// TwinCAT 3 PLC project Untitled1
// ProgramVersion: 3.1.4024.0
// libraries:
//   CmpBitmapPool, * (System)
//   Tc2_ControllerToolbox, * (Beckhoff Automation GmbH)
//   Tc2_MC2, * (Beckhoff Automation GmbH)
//   Tc2_Standard, * (Beckhoff Automation GmbH)
//   Tc2_System, * (Beckhoff Automation GmbH)
//   Tc2_Utilities, * (Beckhoff Automation GmbH)
//   Tc3_Module, * (Beckhoff Automation GmbH)
//   VisuSymbols,3.5.10.0,System
// project tree:
//   DUTs/Cartesian Space/ ST_CartesianAdditionalParametes.TcDUT, ST_CartesianForces.TcDUT, ST_CartesianPose.TcDUT, ST_CartesianState.TcDUT, ST_CartesianTarget.TcDUT, ST_CartesianVelocity.TcDUT
//   DUTs/ En_TargetMode.TcDUT, E_CalibrationState.TcDUT, E_ControllerType.TcDUT, E_GameID.TcDUT, E_Language.TcDUT, E_MainState.TcDUT, E_RehabMode.TcDUT, ST_HomingResult.TcDUT, ST_TherapyConfig.TcDUT
//   DUTs/Joint Space/ ST_JointPose.TcDUT, ST_JointState.TcDUT, ST_JointTarget.TcDUT, ST_JointTorque.TcDUT, ST_JointVelocity.TcDUT
//   / GlobalTextList.TcGTLO, PlcTask.TcTTO, Visualization Manager.TcVMO (not stored)
//   GVLs/ GVL_ConstantCoefficent.TcGVL, GVL_AbsoluteEncoders.TcGVL, GVL_Axes.TcGVL, GVL_Current.TcGVL, GVL_EndeffectorPosition.TcGVL, GVL_ForceTorqueSensor.TcGVL, GVL_GamePong.TcGVL, GVL_HMI.TcGVL, GVL_HomingResult.TcGVL, GVL_MessageStaus.TcGVL, GVL_MicroSwitch.TcGVL, GVL_RobotData.TcGVL, GVL_StatusAxes.TcGVL, GVL_TargetPoints.TcGVL, GVL_Torque.TcGVL
//   POUs/Crazy Car/ FB_CrazyCarGame.TcPOU, ST_CrazyCarToUnity.TcDUT, ST_UnityToCrazyCar.TcDUT
//   POUs/ FB_AdmittanceController.TcPOU, FB_DoHoming.TcPOU, FB_DriveInterface.TcPOU, FB_DynamicsCompensator.TcPOU, FB_ForceController.TcPOU, FB_ForceTorqueSensor.TcPOU, FB_ImpedanceController.TcPOU, FB_LanguageManager.TcPOU, FB_LaunchGame.TcPOU, FB_RobotIsActive.TcPOU, FB_StartGame.TcPOU, FB_SwitchOpMode.TcPOU, FB_TherapyManager.TcPOU, FB_ThreeAxisSafety.TcPOU, FB_RobotKinematics.TcPOU, HardwareWallCheck.TcPOU, MAIN.TcPOU, FB_JointStateReader.TcPOU, FB_VirtuallWall.TcPOU, StopAllMotion.TcPOU
//   POUs/Firrfly Game/ FB_FireflyGame.TcPOU, ST_FireflyFromUnity.TcDUT, ST_FireflyToUnity.TcDUT
//   POUs/HMI_FunBlock/ FB_HMI_Monitoring.TcPOU, FB_HMI_TherapyConfiguration.TcPOU, FB_UserSecuring.TcPOU, MicroswitchCheck.TcPOU
//   POUs/PeelerGame/ ST_PeelerFromUnity.TcDUT, FB_PeelingGame.TcPOU, ST_PeelerToUnity.TcDUT
//   POUs/Sorter Game/ FB_SorterGame.TcPOU, ST_SorterToUnity.TcDUT, ST_UnityToSorter.TcDUT
//   VISUs/ ImagePool.TcIPO (not stored), Screen2.TcVIS, Visualization.TcVIS
// real-time tasks:
//   TASK PlcTask: cycle T#10ms, priority 20, ADS port 350
//   TASK VISU_TASK1: cycle T#200000us, priority 1, ADS port 352
// motion (NC):
//   TASK NC-Task 1 SAF: cycle T#1ms, priority 4, ADS port 501
//   TASK NC-Task 1 SVB: cycle T#1ms, priority 6, ADS port 511
//   AXIS Motor-A (id 1)
//     Velo: Maximum=80
//     OtherSettings: AllowMotionCmdToSlave=true
//     encoder EncType=19
//       EncPara: MaxCount=#xffffffff
//         TimeComp: TimeCompMode=1
//     drive DrvType=16
//       DrvPara: MaxCount=#xffffffff, DriveControlDWord=#x00020000
//         Analog: TorqueSetpointScale=10, ScaleFactorActTorque=0.1
//         TimeComp: TaskDelayCycles=1
//     controller CtrType=1
//       CtrPara: PriorControlFactor=1
//         PosDiffControl: Enable=false
//         Observer: BandWidth=20
//   AXIS Motor-B (id 3)
//     Velo: Maximum=80
//     OtherSettings: AllowMotionCmdToSlave=true
//     encoder EncType=19
//       EncPara: MaxCount=#xffffffff
//         TimeComp: TimeCompMode=1
//     drive DrvType=16
//       DrvPara: MaxCount=#xffffffff, DriveControlDWord=#x00020000
//         Analog: TorqueSetpointScale=10, ScaleFactorActTorque=0.1
//         TimeComp: TaskDelayCycles=1
//     controller CtrType=1
//       CtrPara: PriorControlFactor=1
//         PosDiffControl: Enable=false, Range=20
//         Observer: BandWidth=20
//   AXIS Motor-C (id 2)
//     Velo: Maximum=80
//     OtherSettings: AllowMotionCmdToSlave=true
//     encoder EncType=19
//       EncPara: MaxCount=#xffffffff
//         TimeComp: TimeCompMode=1
//     drive DrvType=16
//       DrvPara: MaxCount=#xffffffff, DriveControlDWord=#x00020000
//         Analog: TorqueSetpointScale=10, ScaleFactorActTorque=0.1
//         TimeComp: TaskDelayCycles=1
//     controller CtrType=1
//       CtrPara: PriorControlFactor=1
//         PosDiffControl: Enable=false
//         Observer: BandWidth=20
// I/O:
//   DEVICE Device 3 (EtherCAT), AmsNetId 10.4.37.185.4.1
//     Motor-A [EPOS4 Module 50/8 EtherCAT]
//       modules: Module 1 (CSP Mode)
//     Motor-B [EPOS4 Module 50/8 EtherCAT]
//       modules: Module 1 (CSP Mode)
//     Motor-C [EPOS4 Module 50/8 EtherCAT]
//       modules: Module 1 (CSP Mode)
//     Box 7 (RFT_EC02) [RFT_EC02]
// variable links:
//   NC-Task 1 SAF/Axes/Motor-A <-> Device 3 (EtherCAT)/Motor-A
//     Drive/Inputs/In/nDataIn3[0] <-> Module 1 (CSP Mode)/CSP Inputs/Torque actual value
//     Drive/Inputs/In/nDcOutputTime <-> InfoData/DcOutputShift
//     Drive/Inputs/In/nState1 <-> Module 1 (CSP Mode)/CSP Inputs/Statusword
//     Drive/Inputs/In/nState2 <-> Module 1 (CSP Mode)/CSP Inputs/Statusword @bit 8
//     Drive/Inputs/In/nState4 @bit 1 <-> WcState/InputToggle
//     Drive/Inputs/In/nState4 <-> WcState/WcState
//     Drive/Inputs/In/nState5 <-> Module 1 (CSP Mode)/CSP Inputs/Mode of operation display
//     Drive/Outputs/Out/nCtrl1 <-> Module 1 (CSP Mode)/CSP Outputs/Controlword
//     Drive/Outputs/Out/nCtrl2 <-> Module 1 (CSP Mode)/CSP Outputs/Controlword @bit 8
//     Drive/Outputs/Out/nCtrl5 <-> Module 1 (CSP Mode)/CSP Outputs/Mode of operation
//     Drive/Outputs/Out/nDataOut1 <-> Module 1 (CSP Mode)/CSP Outputs/Target position
//     Drive/Outputs/Out/nDataOut2 <-> Module 1 (CSP Mode)/CSP Outputs/Target velocity
//     Drive/Outputs/Out/nDataOut3[0] <-> Module 1 (CSP Mode)/CSP Outputs/Torque offset
//     Drive/Outputs/Out/nDataOut4[0] <-> Module 1 (CSP Mode)/CSP Outputs/Target torque
//     Enc/Inputs/In/nDataIn1 <-> Module 1 (CSP Mode)/CSP Inputs/Position actual value
//     Enc/Inputs/In/nDataIn7 <-> Module 1 (CSP Mode)/CSP Inputs/Velocity actual value
//     Enc/Inputs/In/nDcInputTime <-> InfoData/DcInputShift
//     Enc/Inputs/In/nState4 @bit 1 <-> WcState/InputToggle
//     Enc/Inputs/In/nState4 <-> WcState/WcState
//   NC-Task 1 SAF/Axes/Motor-B <-> Device 3 (EtherCAT)/Motor-B
//     Drive/Inputs/In/nDataIn3[0] <-> Module 1 (CSP Mode)/CSP Inputs/Torque actual value
//     Drive/Inputs/In/nDcOutputTime <-> InfoData/DcOutputShift
//     Drive/Inputs/In/nState1 <-> Module 1 (CSP Mode)/CSP Inputs/Statusword
//     Drive/Inputs/In/nState2 <-> Module 1 (CSP Mode)/CSP Inputs/Statusword @bit 8
//     Drive/Inputs/In/nState4 @bit 1 <-> WcState/InputToggle
//     Drive/Inputs/In/nState4 <-> WcState/WcState
//     Drive/Inputs/In/nState5 <-> Module 1 (CSP Mode)/CSP Inputs/Mode of operation display
//     Drive/Outputs/Out/nCtrl1 <-> Module 1 (CSP Mode)/CSP Outputs/Controlword
//     Drive/Outputs/Out/nCtrl2 <-> Module 1 (CSP Mode)/CSP Outputs/Controlword @bit 8
//     Drive/Outputs/Out/nCtrl5 <-> Module 1 (CSP Mode)/CSP Outputs/Mode of operation
//     Drive/Outputs/Out/nDataOut1 <-> Module 1 (CSP Mode)/CSP Outputs/Target position
//     Drive/Outputs/Out/nDataOut2 <-> Module 1 (CSP Mode)/CSP Outputs/Target velocity
//     Drive/Outputs/Out/nDataOut3[0] <-> Module 1 (CSP Mode)/CSP Outputs/Torque offset
//     Drive/Outputs/Out/nDataOut4[0] <-> Module 1 (CSP Mode)/CSP Outputs/Target torque
//     Enc/Inputs/In/nDataIn1 <-> Module 1 (CSP Mode)/CSP Inputs/Position actual value
//     Enc/Inputs/In/nDataIn7 <-> Module 1 (CSP Mode)/CSP Inputs/Velocity actual value
//     Enc/Inputs/In/nDcInputTime <-> InfoData/DcInputShift
//     Enc/Inputs/In/nState4 @bit 1 <-> WcState/InputToggle
//     Enc/Inputs/In/nState4 <-> WcState/WcState
//   NC-Task 1 SAF/Axes/Motor-C <-> Device 3 (EtherCAT)/Motor-C
//     Drive/Inputs/In/nDataIn3[0] <-> Module 1 (CSP Mode)/CSP Inputs/Torque actual value
//     Drive/Inputs/In/nDcOutputTime <-> InfoData/DcOutputShift
//     Drive/Inputs/In/nState1 <-> Module 1 (CSP Mode)/CSP Inputs/Statusword
//     Drive/Inputs/In/nState2 <-> Module 1 (CSP Mode)/CSP Inputs/Statusword @bit 8
//     Drive/Inputs/In/nState4 @bit 1 <-> WcState/InputToggle
//     Drive/Inputs/In/nState4 <-> WcState/WcState
//     Drive/Inputs/In/nState5 <-> Module 1 (CSP Mode)/CSP Inputs/Mode of operation display
//     Drive/Outputs/Out/nCtrl1 <-> Module 1 (CSP Mode)/CSP Outputs/Controlword
//     Drive/Outputs/Out/nCtrl2 <-> Module 1 (CSP Mode)/CSP Outputs/Controlword @bit 8
//     Drive/Outputs/Out/nCtrl5 <-> Module 1 (CSP Mode)/CSP Outputs/Mode of operation
//     Drive/Outputs/Out/nDataOut1 <-> Module 1 (CSP Mode)/CSP Outputs/Target position
//     Drive/Outputs/Out/nDataOut2 <-> Module 1 (CSP Mode)/CSP Outputs/Target velocity
//     Drive/Outputs/Out/nDataOut3[0] <-> Module 1 (CSP Mode)/CSP Outputs/Torque offset
//     Drive/Outputs/Out/nDataOut4[0] <-> Module 1 (CSP Mode)/CSP Outputs/Target torque
//     Enc/Inputs/In/nDataIn1 <-> Module 1 (CSP Mode)/CSP Inputs/Position actual value
//     Enc/Inputs/In/nDataIn7 <-> Module 1 (CSP Mode)/CSP Inputs/Velocity actual value
//     Enc/Inputs/In/nDcInputTime <-> InfoData/DcInputShift
//     Enc/Inputs/In/nState4 @bit 1 <-> WcState/InputToggle
//     Enc/Inputs/In/nState4 <-> WcState/WcState
//   Untitled1/Untitled1 Instance <-> Device 3 (EtherCAT)/Box 7 (RFT_EC02)
//     PlcTask Inputs/GVL_ForceTorqueSensor.RawFx <-> IN_GENERIC process data mapping/Raw_Fx
//     PlcTask Inputs/GVL_ForceTorqueSensor.RawFy <-> IN_GENERIC process data mapping/Raw_Fy
//     PlcTask Inputs/GVL_ForceTorqueSensor.RawFz <-> IN_GENERIC process data mapping/Raw_Fz
//     PlcTask Inputs/GVL_ForceTorqueSensor.RawMx <-> IN_GENERIC process data mapping/Raw_Tx
//     PlcTask Inputs/GVL_ForceTorqueSensor.RawMy <-> IN_GENERIC process data mapping/Raw_Ty
//     PlcTask Inputs/GVL_ForceTorqueSensor.RawMz <-> IN_GENERIC process data mapping/Raw_Tz
//     PlcTask Outputs/GVL_ForceTorqueSensor.ConfigParameter <-> OUT_GENERIC process data mapping/ConfigParam_1
//   Untitled1/Untitled1 Instance <-> Device 3 (EtherCAT)/Motor-A
//     PlcTask Inputs/GVL_AbsoluteEncoders.AbsoluteBetaPosition <-> Module 1 (CSP Mode)/CSP Inputs/Position actual value sensor 2
//     PlcTask Inputs/GVL_Current.MotorCurrentM1_mA <-> Module 1 (CSP Mode)/CSP Inputs/Current actual value averaged
//     PlcTask Inputs/GVL_MicroSwitch.dwMicroSwitchDriverA <-> Module 1 (CSP Mode)/CSP Inputs/Digital inputs
//   Untitled1/Untitled1 Instance <-> Device 3 (EtherCAT)/Motor-B
//     PlcTask Inputs/GVL_AbsoluteEncoders.AbsoluteLinearPosition <-> Module 1 (CSP Mode)/CSP Inputs/Position actual value sensor 2
//     PlcTask Inputs/GVL_Current.MotorCurrentM2_mA <-> Module 1 (CSP Mode)/CSP Inputs/Current actual value averaged
//     PlcTask Inputs/GVL_MicroSwitch.dwMicroSwitchDriverB <-> Module 1 (CSP Mode)/CSP Inputs/Digital inputs
//   Untitled1/Untitled1 Instance <-> Device 3 (EtherCAT)/Motor-C
//     PlcTask Inputs/GVL_AbsoluteEncoders.AbsoluteTetaPosition <-> Module 1 (CSP Mode)/CSP Inputs/Position actual value sensor 2
//     PlcTask Inputs/GVL_Current.MotorCurrentM3_mA <-> Module 1 (CSP Mode)/CSP Inputs/Current actual value averaged
//   Untitled1/Untitled1 Instance <-> NC-Task 1 SAF/Axes/Motor-A
//     PlcTask Inputs/GVL_Axes.Axis1.NcToPlc <-> Outputs/ToPlc
//     PlcTask Inputs/GVL_Torque.TorqueM1_Act <-> Outputs/ToPlc/ActTorque
//     PlcTask Outputs/GVL_Axes.Axis1.PlcToNc <-> Inputs/FromPlc
//   Untitled1/Untitled1 Instance <-> NC-Task 1 SAF/Axes/Motor-B
//     PlcTask Inputs/GVL_Axes.Axis2.NcToPlc <-> Outputs/ToPlc
//     PlcTask Inputs/GVL_Torque.TorqueM2_Act <-> Outputs/ToPlc/ActTorque
//     PlcTask Outputs/GVL_Axes.Axis2.PlcToNc <-> Inputs/FromPlc
//   Untitled1/Untitled1 Instance <-> NC-Task 1 SAF/Axes/Motor-C
//     PlcTask Inputs/GVL_Axes.Axis3.NcToPlc <-> Outputs/ToPlc
//     PlcTask Inputs/GVL_Torque.TorqueM3_Act <-> Outputs/ToPlc/ActTorque
//     PlcTask Outputs/GVL_Axes.Axis3.PlcToNc <-> Inputs/FromPlc

CONFIGURATION Untitled1
    RESOURCE PLC ON TwinCAT3
        TASK PlcTask(INTERVAL := T#10ms, PRIORITY := 20);
        PROGRAM MAIN WITH PlcTask : MAIN;
    END_RESOURCE
END_CONFIGURATION

// ---- DUTs/Cartesian Space/ST_CartesianAdditionalParametes.TcDUT
TYPE ST_CartesianAdditionalParametes :
STRUCT
	BetaIncremental : LREAL;
	RIncremental : LREAL;
	X_Dir_Abs :LREAL;
	Y_Dir_Abs :LREAL;
	WristAngle_Abs : LREAL;

END_STRUCT
END_TYPE

// ---- DUTs/Cartesian Space/ST_CartesianForces.TcDUT
TYPE ST_CartesianForces :
STRUCT
	Fx     : LREAL; // Linear force along X (N)
    Fy     : LREAL; // Linear force along Y (N)
    Mtheta : LREAL; // Moment/Torque around Theta wrist axis (Nm)
END_STRUCT
END_TYPE

// ---- DUTs/Cartesian Space/ST_CartesianPose.TcDUT
TYPE ST_CartesianPose :
STRUCT
	X     : LREAL; // X position (mm)
    Y     : LREAL; // Y position (mm)
    Theta : LREAL; // Wrist angle (deg / rad)
END_STRUCT
END_TYPE

// ---- DUTs/Cartesian Space/ST_CartesianState.TcDUT
TYPE ST_CartesianState :
STRUCT
	Position : ST_CartesianPose;     // Contains X, Y, Theta
    Velocity : ST_CartesianVelocity; // Contains Vx, Vy, Vtheta
	Force    : ST_CartesianForces;    // Contains Fx, Fy, Mtheta
END_STRUCT
END_TYPE

// ---- DUTs/Cartesian Space/ST_CartesianTarget.TcDUT
TYPE ST_CartesianTarget :
STRUCT
	Position : ST_CartesianPose;     // Game target position
    Velocity : ST_CartesianVelocity; // Feedforward target velocity
    Force    : ST_CartesianForces;    // Force setpoint (e.g. 0 N for admittance)
END_STRUCT
END_TYPE

// ---- DUTs/Cartesian Space/ST_CartesianVelocity.TcDUT
TYPE ST_CartesianVelocity :
STRUCT
	Vx     : LREAL; // Linear velocity along X (mm/s or m/s)
    Vy     : LREAL; // Linear velocity along Y (mm/s or m/s)
    Vtheta : LREAL; // Angular velocity around Theta (deg/s or rad/s)
END_STRUCT
END_TYPE

// ---- DUTs/En_TargetMode.TcDUT
{attribute 'qualified_only'}
{attribute 'strict'}
TYPE En_TargetMode :
(
	eCSP := 4,   // Cyclic Synchronous Position
    eCSV := 2,   // Cyclic Synchronous Velocity
    eCST := 1   // Cyclic Synchronous Torque
);
END_TYPE

// ---- DUTs/E_CalibrationState.TcDUT
{attribute 'qualified_only'}
{attribute 'strict'}
TYPE E_CalibrationState :
(
	INIT,
    SET_FILTER,
    START,
    WaitingforCalibrationButton,
    ZEROING,
    RUNNING
);
END_TYPE

// ---- DUTs/E_ControllerType.TcDUT
{attribute 'qualified_only'}
{attribute 'strict'}
TYPE E_ControllerType :
(
    ControlNone         := 0,

    ControlPosition     := 1,

    ControlVelocity     := 2,

    ControlTorque       := 3,

    ControlForce        := 4,

    ControlImpedance    := 5,

    ControlAdmittance   := 6,

    ControlHybrid       := 7,

    ControlCustom       := 8
);
END_TYPE

// ---- DUTs/E_GameID.TcDUT
{attribute 'qualified_only'}
{attribute 'strict'}
TYPE E_GameID :
(
    NONE        := 0,
    PONG        := 1,
    PEELING     := 2,
    GOLD_MINER  := 3,
    BALLOON     := 4,
    SNOW_WIPER  := 5,
    SORTER      := 6,
    FLOWER      := 7,
    CRAZY_CAR   := 8
);
END_TYPE

// ---- DUTs/E_Language.TcDUT
{attribute 'qualified_only'}
{attribute 'strict'}
TYPE E_Language :
(
	EN,
    FR
);
END_TYPE

// ---- DUTs/E_MainState.TcDUT
{attribute 'qualified_only'}
{attribute 'strict'}
TYPE E_MainState :
(
	Init                := 0,
    Homing              := 10,
    ClearNCErrors       := 20,
    ChangingDriverMode        := 30,
    Standby             := 40,  // NEW: Motors are ON, holding position, waiting for HMI start
    RunningTherapy      := 50,  // NEW: The robot is actively doing rehab
    Fault               := 99
);
END_TYPE

// ---- DUTs/E_RehabMode.TcDUT
{attribute 'qualified_only'}
{attribute 'strict'}
TYPE E_RehabMode :
(
	ModeIdle              := 0, // Safety default: system is ready but therapy is not active
    ModePassive           := 1, // Robot moves a completely relaxed patient rigidly along a path
    ModeActiveFree        := 2, // Robot is totally transparent; patient moves freely without resistance
    ModeActiveAssistive   := 3, // Robot provides assistive forces to help the patient reach the target
    ModeActiveResistive   := 4, // Robot pushes against the patient to build muscle strength
    ModePerturbation      := 5, // Robot applies sudden, unexpected forces to train patient reflexes
    ModeAssessment        := 6  // Robot measures patient capability passively without providing assistance
);
END_TYPE

// ---- DUTs/Joint Space/ST_JointPose.TcDUT
TYPE ST_JointPose :
STRUCT
	q1 : LREAL;
    q2 : LREAL;
    q3 : LREAL;
END_STRUCT
END_TYPE

// ---- DUTs/Joint Space/ST_JointState.TcDUT
TYPE ST_JointState :
STRUCT
	Position : ST_JointPose; // Current joint angles (J1, J2, J3)
    Velocity : ST_JointVelocity; // Current joint speeds (J1, J2, J3)
    Torque   : ST_JointTorque; // Measured motor torques (J1, J2, J3)
END_STRUCT
END_TYPE

// ---- DUTs/Joint Space/ST_JointTarget.TcDUT
TYPE ST_JointTarget :
STRUCT
	Position : ST_JointPose; // Commanded joint angles
    Velocity : ST_JointVelocity; // Commanded joint speeds
    Torque   : ST_JointTorque; // Calculated motor torques (T1, T2, T3)
END_STRUCT
END_TYPE

// ---- DUTs/Joint Space/ST_JointTorque.TcDUT
TYPE ST_JointTorque :
STRUCT
	M1 : LREAL;
    M2 : LREAL;
    M3 : LREAL;
END_STRUCT
END_TYPE

// ---- DUTs/Joint Space/ST_JointVelocity.TcDUT
TYPE ST_JointVelocity :
STRUCT
	q1_dot : LREAL; // dq1 / dt
    q2_dot : LREAL; // dq2 / dt
    q3_dot : LREAL; // dq3 / dt
END_STRUCT
END_TYPE

// ---- DUTs/ST_HomingResult.TcDUT
TYPE ST_HomingResult :
STRUCT
	HomePos_Beta  : LREAL;   (* joint angle/position after homing *)
    HomePos_Theta  : LREAL;
    HomePos_R  : LREAL;
END_STRUCT
END_TYPE

// ---- DUTs/ST_TherapyConfig.TcDUT
TYPE ST_TherapyConfig :
STRUCT
	// 1. Core Selections
    TherapyMode          : E_RehabMode;
    ControllerType       : E_ControllerType;
    
    // 2. Feature Flags
    FeatureInertiaComp   : BOOL;  
    FeatureFrictionComp  : BOOL; 
    FeatureVirtualWall   : BOOL; 
	
//    FeatureDataLogger    : BOOL; 
    
    // 3. Global Safety Limits (Apply to ALL controllers)
    GlobalForceLimit     : LREAL := 50 ; // Maximum safe force allowed
    GlobalVelocityLimit  : LREAL; // Maximum safe speed allowed (please clarify : is it in Jointspace or Cartesian space)
	
	Stiffness_K         : LREAL; // Virtual spring stiffness for Impedance
    Damping_D           : LREAL; // Virtual friction/viscosity for Impedance
    Mass_M              : LREAL; // Virtual mass for Admittance
END_STRUCT
END_TYPE

// ---- POUs/Crazy Car/ST_CrazyCarToUnity.TcDUT
TYPE ST_CrazyCarToUnity :
STRUCT
	fY           : REAL;   // gas, Y position 0..100 %
    fWristAngle  : REAL;   // wrist angle, degrees, 0 = home
    GameIsActive : BOOL;
END_STRUCT
END_TYPE

// ---- POUs/Crazy Car/ST_UnityToCrazyCar.TcDUT
TYPE ST_UnityToCrazyCar  :
STRUCT
	bGameClosed : BOOL;   // TRUE = Unity game closed
    nGameStatus : INT;    // 0 = menu/popup, 1 = Taxi, 2 = Van, 3 = Truck
END_STRUCT
END_TYPE

// ---- POUs/Firrfly Game/ST_FireflyFromUnity.TcDUT
{attribute 'pack_mode' := '1'}
TYPE ST_FireflyFromUnity :
STRUCT
    nGameStatus  : INT;    // 0 = menu/results, 1/2/3 = playing Level 1/2/3, 4 = paused
    bExitPressed : BOOL;   // TRUE for ~0.2 s when an Exit button is pressed, then FALSE
    bWrongFlower : BOOL;   // TRUE for ~0.2 s each time a wrong flower is selected, then FALSE
END_STRUCT
END_TYPE

// ---- POUs/Firrfly Game/ST_FireflyToUnity.TcDUT
TYPE ST_FireflyToUnity :
STRUCT
    fX : REAL;   // -100..+100 %, 0 = home (middle of the scene), +100 = right edge of the garden
    fY : REAL;   // -100..+100 %, 0 = home (middle of the scene), +100 = top edge (robot forward)
END_STRUCT
END_TYPE

// ---- POUs/PeelerGame/ST_PeelerFromUnity.TcDUT
{attribute 'pack_mode' := '1'}
TYPE ST_PeelerFromUnity :
STRUCT
	bInContact    : BOOL;    // Fruit collision state
    nObjectType   : INT;     // 1 = Kiwi, 2 = Orange, 3 = Pineapple
    bGameFinished : BOOL;    // TRUE when the user clicks the Close button in Unity
END_STRUCT
END_TYPE

// ---- POUs/PeelerGame/ST_PeelerToUnity.TcDUT
TYPE ST_PeelerToUnity :
STRUCT
	fY          : REAL;    // Y position (0 - 100%)
	GameIsActive : BOOL;
   

END_STRUCT
END_TYPE

// ---- POUs/Sorter Game/ST_SorterToUnity.TcDUT
TYPE ST_SorterToUnity :
STRUCT
    fX           : REAL;    // X position 0–100%
    GameIsActive : BOOL;
END_STRUCT
END_TYPE

// ---- POUs/Sorter Game/ST_UnityToSorter.TcDUT
TYPE ST_UnityToSorter :
STRUCT
	bGameClosed : BOOL;   // TRUE = Unity game closed
    nGameStatus : INT;    // 0 = not playing, 1 = light, 2 = medium, 3 = heavy
END_STRUCT
END_TYPE

// ---- GVLs/GVL_ConstantCoefficent.TcGVL
{attribute 'qualified_only'}
// These number is checked two times, the error between Absolute and Incremental Encoder is under 1% that is acceptable
// Root of error is related to timing belt 


VAR_GLOBAL
	K2: LREAL :=24.40;  // calculate with result of absolute encoder
	
	K3: LREAL :=219.726; // calculate with result of absolute encoder
	K1: LREAL := 9.97; // calculate with result of absolute encoder
	
END_VAR

// ---- GVLs/GVL_AbsoluteEncoders.TcGVL
{attribute 'qualified_only'}
VAR_GLOBAL
	AbsoluteBetaPosition AT %I* : DINT;
	AbsoluteLinearPosition AT %I* : DINT;
	AbsoluteTetaPosition AT %I* : DINT;
END_VAR

// ---- GVLs/GVL_Axes.TcGVL
{attribute 'qualified_only'}
VAR_GLOBAL
	Axis1 : AXIS_REF;
	Axis2 : AXIS_REF;
	Axis3 : AXIS_REF;
END_VAR

// ---- GVLs/GVL_Current.TcGVL
{attribute 'qualified_only'}
VAR_GLOBAL
	MotorCurrentM1_mA AT %I* : DINT; // PDO value from EPOS4 [mA]
	MotorCurrentM2_mA AT %I* : DINT;
	MotorCurrentM3_mA AT %I* : DINT;
	MotorCurrentM1_A : LREAL;  // // Converted current [A]
	MotorCurrentM2_A : LREAL;
	MotorCurrentM3_A : LREAL;
	
END_VAR

// ---- GVLs/GVL_EndeffectorPosition.TcGVL
{attribute 'qualified_only'}
VAR_GLOBAL
	WristAngle : LREAL;
	X_Dir : LREAL;
	Y_Dir : LREAL;
	R_Dir : LREAL;
	Beta : LREAL;
	
	X_Dir_Abs: LREAL;
	Y_Dir_Abs: LREAL;
	R_Dir_Abs: LREAL;
	BetaFromAbsolute : LREAL;
	WristAngle_Abs: LREAL;
	
END_VAR

// ---- GVLs/GVL_ForceTorqueSensor.TcGVL
{attribute 'qualified_only'}
VAR_GLOBAL
	ConfigParameter AT %Q* : DWORD;
	RawFx AT %I* : INT;
	RawFy AT %I* : INT;
	RawFz AT %I* : INT;
	RawMx AT %I* : INT;
	RawMy AT %I* : INT;
	RawMz AT %I* : INT;
	
	//
	Fx_ActFTS : LREAL;    // N
	Fy_ActFTS : LREAL;
	Mz_ActFTS : LREAL;    //N.M
	
END_VAR

// ---- GVLs/GVL_GamePong.TcGVL
{attribute 'qualified_only'}
VAR_GLOBAL
	// Robot Position for Unity (0-100)
    MyRobotY : REAL ;
END_VAR

// ---- GVLs/GVL_HMI.TcGVL
{attribute 'qualified_only'}
VAR_GLOBAL
	


	
	bLaunchGameSpongCmd : BOOL := FALSE;
	bLaunchGamePeelerCmd : BOOL := FALSE;
	bLaunchGameGoldMiner : BOOL := FALSE;
	bLaunchGameBalloonAssesment : BOOL := FALSE;
	bLaunchGameSnowWiper : BOOL := FALSE;
	bLaunchGameSorter : BOOL := FALSE;
	bLaunchGameFlower : BOOL := FALSE;
	bLaunchGameCrazyCar : BOOL := FALSE;
	
	
	
	
	
	// MicroSwitch Check
	CheckMicroswitchLinearMin : BOOL := FALSE;
	CheckMicroswitchLinearMax : BOOL := FALSE;
	CheckMicroswitchRotationLeft : BOOL := FALSE;
	CheckMicroswitchRotationRight : BOOL := FALSE;
	CheckMicroswitchWristLeft : BOOL := FALSE;
	CheckMicroswitchWristRight : BOOL := FALSE;
	
	HardwareLimitisActived : BOOL := FALSE;
	
	
			// HMIHardwareMicroSwitch Check for activation
	
	HwCheckMicroswitchLinearMin : BOOL := FALSE;
	HwCheckMicroswitchLinearMax : BOOL := FALSE;
	HwCheckMicroswitchRotationLeft : BOOL := FALSE;
	HwCheckMicroswitchRotationRight : BOOL := FALSE;
	HwCheckMicroswitchWristLeft : BOOL := FALSE;
	HwCheckMicroswitchWristRight : BOOL := FALSE;
	
	// TurningonPageinHMI when hardwarelimit Activated
	
	
	ContinueToHoming : BOOL := FALSE;
	StartTherapy: BOOL;
	StartRobot_HMI : BOOL;
	StartHomingDisable_HMI : BOOL := TRUE;
	ContinueToSensorCalibrationDisable_HMI : BOOL := FALSE;
	Homingprogress : UINT;
	StartCalibrationButton : BOOL := FALSE;
	UserSecuringButton_HMI : BOOL := FALSE;
	Fx_HMI: LREAL;
	Fy_HMI: LREAL;
	Mz_HMI: LREAL;
	SecuringPage : INT :=1 ;
	
	
	// User Securing
	check1 : BOOL := FALSE;
	check2 : BOOL := FALSE;
	check3 : BOOL := FALSE;
	check4 : BOOL := FALSE;
	check5 : BOOL := FALSE;
	check6 : BOOL := FALSE;
	ContinueTOWorkspaceLimits : BOOL := FALSE;
	MainPageButtonEnableDisable : BOOL :=FALSE;
	EmergencyStopIsOnHardware : BOOL := FALSE;
	EmergencyStopIsOnSoftware : BOOL := FALSE;
	HomingError : BOOL := FALSE;
	CurrentTherapyConfig : ST_TherapyConfig;
	Virtuallwall : BOOL;
	VirtualWallContact : BOOL;
	EndeffectorPositionPixcelUnit_X : INT;
	EndeffectorPositionPixcelUnit_Y : INT;
	EndeffectorPositionPixcelUnit_Theta : LREAL;
	
PolygonPoints : STRING(255);

  // Variable related to Workspace

  // Hardware Limit Switches
   

    bRotationLeftLimit        : BOOL;
    bRotationRightLimit       : BOOL;

    bLinearMaxLimit           : BOOL;
    bLinearMinLimit           : BOOL;

    bWristRightLimit          : BOOL;
    bWristLeftLimit           : BOOL;
	
	
	EableVirtuallWall_Planar : BOOL;
	EnableWristWall : BOOL;
	// PLanar Button

	TopPlanarWall_But : BOOL;
	BottomPlanarWall_But : BOOL;
	RightPlanarWall_But: BOOL;
	LeftPlanarWall_But : BOOL;
	
	SETPlanarWall_But : BOOL;
	
	RightWristWall_But : BOOL;
	LeftWristWall_But : BOOL;
	SETWristWall_But : BOOL;
	







// Therapy Configuration
	
	    // Global safety limits
    MaxForce : LREAL := 20.0;
    MaxVelocity : LREAL := 50.0;


    // Therapy mode
    TherapyMode : INT := 0;

    bActiveMode : BOOL := FALSE;
    bPassiveMode : BOOL := FALSE;
    bAssistiveMode : BOOL := FALSE;
    bResistiveMode : BOOL := FALSE;
    bGameBasedMode : BOOL := TRUE;


    // Dynamics compensation
    bFrictionCompensation : BOOL := FALSE;
    bInertiaCompensation : BOOL := FALSE;


    // Control type
    ControlType : INT := 0;

    bImpedanceControl : BOOL := TRUE;
    bAdmittanceControl : BOOL := FALSE;


    // Control parameters
    Stiffness : LREAL := 20.5;
    Damping : LREAL := 0.0;
    Mass : LREAL := 0.0;


    // Start therapy
    bStartTherapy : BOOL := FALSE;
	
	
END_VAR

// ---- GVLs/GVL_HomingResult.TcGVL
{attribute 'qualified_only'}
VAR_GLOBAL
	gHoming : ST_HomingResult;
END_VAR

// ---- GVLs/GVL_MessageStaus.TcGVL
{attribute 'qualified_only'}
VAR_GLOBAL
	MessageStaus : STRING(255);	
END_VAR

// ---- GVLs/GVL_MicroSwitch.TcGVL
{attribute 'qualified_only'}
VAR_GLOBAL
	dwMicroSwitchDriverA AT %I* : DWORD;
	dwMicroSwitchDriverB AT %I* : DWORD;
END_VAR

// ---- GVLs/GVL_RobotData.TcGVL
{attribute 'qualified_only'}
VAR_GLOBAL
	Q1_Actual : LREAL;
    Q2_Actual : LREAL;
    Q3_Actual : LREAL;
END_VAR

// ---- GVLs/GVL_StatusAxes.TcGVL
{attribute 'qualified_only'}
VAR_GLOBAL
	ErrorAxis1 	AT %I* : INT;
	ErrorAxis2 	AT %I*: INT;
	ErrorAxis3 	AT %I*: INT;
	//Driver1Status AT %I* : UINT;
	Driver2Status AT %I* : UINT;
	Driver3Status AT %I* : UINT;
	
END_VAR

// ---- GVLs/GVL_TargetPoints.TcGVL
{attribute 'qualified_only'}
VAR_GLOBAL
	Target_A : ARRAY [1..3] OF LREAL := [0.0, 200.0, 0.0];
    Target_B : ARRAY [1..3] OF LREAL := [450.0, 100.0, 30.0];
    Target_C : ARRAY [1..3] OF LREAL := [450.0, -100.0, -30.0];
END_VAR

// ---- GVLs/GVL_Torque.TcGVL
{attribute 'qualified_only'}
VAR_GLOBAL
	TorqueM1_Act AT %I* : LREAL;
	TorqueM2_Act AT %I* : LREAL;
	TorqueM3_Act AT %I* : LREAL;
	TorqueM33_Act : LREAL;
END_VAR

// ---- POUs/MAIN.TcPOU
PROGRAM MAIN
VAR
	
	fbMC_Power1: MC_Power;
	xEnable: BOOL;
	xControlPower: BOOL;
	fbMC_Power2: MC_Power;
	fbMC_Power3: MC_Power;
	fbMC_Reset: MC_Reset;
	fbMC_Reset1: MC_Reset;
	xAxisReset: BOOL;
	fbMC_Reset2: MC_Reset;
	fbMC_Reset3: MC_Reset;
	xMachineReset: BOOL;
	eState: INT := 0;
	// Homming
	HomingDone: BOOL;
	HomingStart: BOOL;
	fbDoHoming : FB_DoHoming;
	bHomingError: BOOL;
	 WaitForStartHoming : TON;
	 rtStartHoming : R_TRIG;
	 HomingProgressTime : TON;
	//Safety
	fbSafety : FB_ThreeAxisSafety;
	fbEmergencyStop : StopAllMotion;
	RobotIsNotSafe: BOOL;
	
	AbsEncDegNutralPos: UDINT;
	
	// READ POSITION
	fbJointReader    : FB_JointStateReader;
	ActualJoints     : ST_JointState;      // Joint feedback (q, q_dot, M)
	ActualCartesian : ST_CartesianState;
	JointDataTransedFromCartesianSpace : ST_JointState;
	CartesianDataTransedFromJointSpace : ST_CartesianState;
	ActualCartesianPose_PERCENTAGE : ST_CartesianPose;
	ActualCartesianAbsolute : ST_CartesianAdditionalParametes;
	AdditionalPose : ST_CartesianAdditionalParametes;
	fbKinematicRobot : FB_RobotKinematics;
	fbReadPosM1 : MC_ReadActualPosition;
	fbReadPosM2 : MC_ReadActualPosition;
	fbReadPosM3 : MC_ReadActualPosition;
	AA: LREAL;
	xDir: LREAL;
	yDir: LREAL;
	theta: LREAL;
	betaAngle : LREAL;
	justfortestrepository : INT;
	EndeffectorVelociybyJacobian : ST_CartesianVelocity;
	
	// visualization
	Point1 : INT;
	
	fbRobotisActive : FB_RobotIsActive;
	
	


// Active Mode
	A_Point : ARRAY [1..3] OF LREAL;  // x, y , and theta (wrist) in A point
	B_Point : ARRAY [1..3] OF LREAL;  // x, y , and theta (wrist) in A point
	C_Point : ARRAY [1..3] OF LREAL;  // x, y , and theta (wrist) in A point
	
	
	OperationalMode : En_TargetMode;
	bExecuteChangingMode : BOOL := FALSE;
	bSwitchopModeDone : BOOL := FALSE;
	fbSwitchMode : FB_SwitchOpMode;
	BActiveMode: BOOL := FALSE;
	ANNModeIsDone : BOOL;
	// Games
	myGameLauncher : FB_LaunchGame;
	eActiveGame : E_GameID;
	
	fbSorterGame : FB_SorterGame;
	fbCrazyCar : FB_CrazyCarGame;
	fbFireflyGame : FB_FireflyGame;

	
	// Force Torque Sensor
	fbForceTorqueSensor : FB_ForceTorqueSensor;
	
	//HMI
	fbMicroswitchCheck : MicroswitchCheck;
	fbUserSecurity : FB_UserSecuring;
	
	StatusOfEmergencyStop: STRING;
	EmergenywasActive: BOOL;
	
	// Rehabilitation mode
	 eMode : E_RehabMode;
	 fbTherapyManager : FB_TherapyManager;
	 
	 fbDriveInterface: FB_DriveInterface;
	 
	TargetJointsextractedfromfbThetapyManger : ST_JointTorque;
	fbHMITemporary : FB_HMI_TherapyConfiguration;
	ERRORIDAxis1: UDINT;
	ERRORIDAxis2: UDINT;
	ERRORIDAxis3: UDINT;
	fbPeelingGame : FB_PeelingGame;
	stGameTargetTorque : ST_JointTorque;
	fbVirtuallWall : FB_VirtuallWall;
	// hardwaresafety
	FirsttimeCheckMicroawitch: BOOL := TRUE;
	CheckingHardwareAcrivation : HardwareWallCheck;
	Hardwaresafetylimit : BOOL;
	
	WallSetPointXandY : ARRAY[1..4, 1..2] OF LREAL;
END_VAR

(* Actuaros Current Status *)
// You can Delete this section 
// This section is implemented Just for checking safety 
GVL_Current.MotorCurrentM1_A :=
    DINT_TO_LREAL(GVL_Current.MotorCurrentM1_mA) / 1000.0;
GVL_Current.MotorCurrentM2_A :=
    DINT_TO_LREAL(GVL_Current.MotorCurrentM2_mA) / 1000.0;
GVL_Current.MotorCurrentM3_A :=
    DINT_TO_LREAL(GVL_Current.MotorCurrentM3_mA) / 1000.0;



//HMI 
fbMicroswitchCheck();
fbUserSecurity();





// Read Status
GVL_Axes.Axis1.ReadStatus();
GVL_Axes.Axis2.ReadStatus();
GVL_Axes.Axis3.ReadStatus();
(*
//Games
myGameLauncher(
    bTrigger    := GVL_HMI.bLaunchGameSpongCmd,
    sExePath    := 'C:\Users\hkhabiri\Desktop\PongV2\RobotGame_BuildV4\Pong.exe', 
    sWorkingDir := 'C:\Users\hkhabiri\Desktop\PongV2\RobotGame_BuildV4\'
	  
);

myGameLauncher(
    bTrigger    := GVL_HMI.bLaunchGamePeelerCmd,
    sExePath    := 'C:\Users\hkhabiri\Desktop\MotivaGames\KIWIexe\First_Project.exe', 
    sWorkingDir := 'C:\Users\hkhabiri\Desktop\MotivaGames\KIWIexe\'
	  
);

*)
// Read Absolute Encoder

//AbsEncDegNutralPos := GVL_AbsoluteEncoder.SSI_Raw32;


// Binding TO HMI Variables
xControlPower := GVL_HMI.StartRobot_HMI;


//EnablefbMC_Power1(
	IF xControlPower THEN
		xEnable := TRUE;
	ELSE
			xEnable := FALSE;
	END_IF
	


// Force-Torque Sensor	
		
	
	fbMC_Power1(
		Axis:= GVL_Axes.Axis1 , 
		
		Enable_Positive:= xEnable , 
		Enable_Negative:= xEnable , 
		Override:= 100.0 );
	fbMC_Power2(
		Axis:= GVL_Axes.Axis2 , 
		
		Enable_Positive:= xEnable , 
		Enable_Negative:= xEnable , 
		Override:= 100.0 );	
	fbMC_Power3(
		Axis:= GVL_Axes.Axis3 , 
		
		Enable_Positive:= xEnable , 
		Enable_Negative:= xEnable , 
		Override:= 100.0  );
		
	IF estate <> 20 THEN 
		fbMC_Power1.Enable:= xEnable;
		fbMC_Power2.Enable:= xEnable;
		fbMC_Power3.Enable:= xEnable;
		
					
	END_IF
	
	IF estate = 20 THEN 
		
	xControlPower:= FALSE; 
	
	END_IF
	
// Reset
	IF xMachineReset THEN
		xAxisReset:= TRUE;
		ELSE
		xAxisReset:= FALSE;
		END_IF
	
(*	fbMC_Reset1(
		Axis:= GVL_Axes.Axis1 , 
		Execute:= xAxisReset AND GVL_Axes.Axis1.Status.Error);
	fbMC_Reset2(
		Axis:= GVL_Axes.Axis2 , 
		Execute:= xAxisReset AND GVL_Axes.Axis2.Status.Error);
	fbMC_Reset3(
		Axis:= GVL_Axes.Axis3 , 
		Execute:= xAxisReset AND GVL_Axes.Axis3.Status.Error); *)

// EmergencyConditionStaus
IF GVL_Axes.Axis1.Status.Error OR GVL_Axes.Axis2.Status.Error OR GVL_Axes.Axis3.Status.Error THEN
	ERRORIDAxis1 := GVL_Axes.Axis1.Status.ErrorID;
	ERRORIDAxis2 := GVL_Axes.Axis2.Status.ErrorID;
	ERRORIDAxis3 := GVL_Axes.Axis3.Status.ErrorID;
	GVL_HMI.EmergencyStopIsOnHardware := TRUE; // YOu can change it if in middle of the work Drivers go to Error
END_IF

IF GVL_HMI.EmergencyStopIsOnSoftware OR GVL_HMI.EmergencyStopIsOnHardware THEN
	eState := E_MainState.Fault;
// fbEmergencyStop ();	
EmergenywasActive := TRUE;

END_IF

IF EmergenywasActive AND NOT GVL_HMI.EmergencyStopIsOnSoftware AND NOT GVL_HMI.EmergencyStopIsOnHardware THEN
eState := E_MainState.Fault;
//fbEmergencyStop ();	
EmergenywasActive := FALSE;
END_IF

// Safety
IF HomingDone THEN
fbSafety(AnyError => RobotIsNotSafe );		
END_IF

//READ PHYSICAL MOTOR HARDWARE
// Updates Joint Positions (q), Velocities (q_dot), and Torques (M)
fbJointReader(
    Axis1      := GVL_Axes.Axis1,
    Axis2      := GVL_Axes.Axis2,
    Axis3      := GVL_Axes.Axis3,
    JointState => ActualJoints
);


fbKinematicRobot( JointData_INPUT:= ActualJoints,
			CartesianData_INPUT := ActualCartesian,
    		JointData_Transed =>  JointDataTransedFromCartesianSpace ,
			CartesianData_Transed => CartesianDataTransedFromJointSpace,
			Cartesian_PERCENTAGE_PoseObtainedFromForwardKinematic => ActualCartesianPose_PERCENTAGE,
			AdditionalPOSE  => AdditionalPose);
			
			
fbHMITemporary(CartesianDataTransedFromJointSpace :=CartesianDataTransedFromJointSpace, WallSetPointXandY=> WallSetPointXandY);
(*
// Reading encoder data
fbReadPosM1(Axis := GVL_Axes.Axis1, Enable := TRUE);
fbReadPosM2(Axis := GVL_Axes.Axis2, Enable := TRUE);
fbReadPosM3(Axis := GVL_Axes.Axis3, Enable := TRUE);
	GVL_RobotData.Q1_Actual := fbReadPosM1.Position;
	GVL_RobotData.Q2_Actual := fbReadPosM2.Position;
	GVL_RobotData.Q3_Actual := fbReadPosM3.Position;
		
// KinematicDATA
fbKinematic(q1:=GVL_RobotData.Q1_Actual, 
				q2:=GVL_RobotData.Q2_Actual,
				q3:=GVL_RobotData.Q3_Actual);	
	
*)
	
// Force-Torque Sensor
fbForceTorqueSensor(CartesianState := ActualCartesian);   // Force-Torque Calibration and Reading


	
	
	
// Robot Operate		
CASE eState OF

E_MainState.Init: (* INIT *)

    HomingDone := FALSE;
    HomingStart := FALSE;

    WaitForStartHoming(
        IN := xControlPower,
        PT := T#0.2S
    );
	IF xControlPower THEN
		GVL_HMI.StartHomingDisable_HMI := FALSE;
	END_IF

    IF WaitForStartHoming.Q THEN
        eState := E_MainState.Homing;
    END_IF


E_MainState.Homing: (* HOMING *)

    WaitForStartHoming(
        IN := FALSE,
        PT := T#2S
    );

    HomingStart := TRUE;
HomingProgressTime (IN :=HomingStart, PT :=T#40S);
GVL_HMI.Homingprogress :=
    DINT_TO_UINT(
        TIME_TO_DINT(HomingProgressTime.ET) * 100 / 40000
    );
    fbDoHoming(
        HStart := HomingStart,
        HM123Done => HomingDone,
        HomingError => bHomingError
    );
	// Display Homing Error on HMI
	IF bHomingError THEN
		GVL_HMI.HomingError := TRUE;
	END_IF
	
	//

    IF HomingDone AND HomingProgressTime.Q THEN
        HomingStart := FALSE;
		GVL_HMI.ContinueToSensorCalibrationDisable_HMI := TRUE;
        eState := E_MainState.ChangingDriverMode;
    END_IF
	
	E_MainState.ChangingDriverMode:  // Changing Driver MODE ; Switch to CST
	 OperationalMode := En_TargetMode.eCST; // Ensure this is defined in your Enum
        fbSwitchMode(TargetMode := OperationalMode, Done => bSwitchopModeDone);
        
        IF bSwitchopModeDone THEN
            bExecuteChangingMode := FALSE;
			fbMC_Power1.Enable := TRUE;
			fbMC_Power2.Enable := TRUE;
			fbMC_Power3.Enable := TRUE;
            eState := E_MainState.RunningTherapy;
			IF  FirsttimeCheckMicroawitch THEN
				GVL_hmi.CheckMicroswitchLinearMax := FALSE;
				GVL_hmi.CheckMicroswitchLinearMin := FALSE;
				GVL_hmi.CheckMicroswitchRotationLeft := FALSE;
				GVL_hmi.CheckMicroswitchRotationRight := FALSE;
				GVL_HMI.CheckMicroswitchWristLeft := FALSE;
				GVL_HMI.CheckMicroswitchWristRight := FALSE;
				FirsttimeCheckMicroawitch := FALSE;

			END_IF
        ELSE
            bExecuteChangingMode := TRUE;
        END_IF
	

    E_MainState.RunningTherapy: (* RUN therapy --- CORE!*)
	

	 	
  // Activation of Hardware limit

CheckingHardwareAcrivation(HardwareActive => Hardwaresafetylimit);

IF Hardwaresafetylimit THEN
	
	GVL_HMI.HardwareLimitisActived := TRUE;
	eState :=E_MainState.Fault;
	
	
END_IF


 

   
// 2. The Robot is active! Feed the Config and Data to the Manager
            fbTherapyManager(
                Enable         := TRUE,
                Config         := GVL_HMI.CurrentTherapyConfig, // Passes your entire STRUCT!
				WallSetPointXandY := WallSetPointXandY,
				SimpleJointTorqueObtainedFromGames := stGameTargetTorque,
				ActualCartesian := CartesianDataTransedFromJointSpace,
				fbKinematics := fbKinematicRobot,
				TargetJointsTorque => TargetJointsextractedfromfbThetapyManger 
           );
			
			fbDriveInterface( TorqueSetpoints := TargetJointsextractedfromfbThetapyManger,Config := GVL_HMI.CurrentTherapyConfig);
      
 // GAME
 myGameLauncher(
    bLaunchSpong     := GVL_HMI.bLaunchGameSpongCmd,
    bLaunchPeeler    := GVL_HMI.bLaunchGamePeelerCmd,
    bLaunchGoldMiner := GVL_HMI.bLaunchGameGoldMiner,
    bLaunchBalloon   := GVL_HMI.bLaunchGameBalloonAssesment,
    bLaunchSnowWiper := GVL_HMI.bLaunchGameSnowWiper,
    bLaunchSorter    := GVL_HMI.bLaunchGameSorter,
    bLaunchFlower    := GVL_HMI.bLaunchGameFlower,
    bLaunchCrazyCar  := GVL_HMI.bLaunchGameCrazyCar,
    eActiveGame      => eActiveGame
);

fbPeelingGame(
    bEnable                   := (eActiveGame = E_GameID.PEELING),
    stCartesianPosePercentage := ActualCartesianPose_PERCENTAGE,   // From Kinematics
    CartesianForcefY       := ActualCartesian.Force.Fy,      // From Kinematics
    CartesianVy := CartesianDataTransedFromJointSpace.Velocity.Vy
	
  //  stJointTargetTorque       => stGameTargetTorque     // Output torque from game
);

// Sorter Game

fbSorterGame(
    bEnable                    := (eActiveGame = E_GameID.SORTER),
    stCartesianPosePercentage  := ActualCartesianPose_PERCENTAGE,                     // From Kinematics
    CartesianForcefX           := ActualCartesian.Force.Fx,                           // From Force Sensor
    CartesianVx                := CartesianDataTransedFromJointSpace.Velocity.Vx     // From Kinematics
    
  //  stJointTargetTorque        => stGameTargetTorque                                  // Output torque from game
);

// Crazy Car Game
fbCrazyCar(
    bEnable                   := (eActiveGame = E_GameID.CRAZY_CAR),
    stCartesianPosePercentage := ActualCartesianPose_PERCENTAGE,                         // Y 0..100 %
    fWristAngleDeg            := CartesianDataTransedFromJointSpace.Position.Theta,      // degrees
    CartesianVtheta           := CartesianDataTransedFromJointSpace.Velocity.Vtheta,
    CartesianMtheta           := ActualCartesian.Force.Mtheta                           // from force sensor
	//stJointTargetTorque       => stGameTargetTorque     // Output torque from game
);	


// Firefly Garden
fbFireflyGame(
    bEnable                    := (eActiveGame = E_GameID.FLOWER),
    stCartesianPosePercentage  := ActualCartesianPose_PERCENTAGE        // From Kinematics (X and Y)
//  stJointTargetTorque        => stGameTargetTorque                    // Output torque from game (always 0: motion only)
);	
			
stGameTargetTorque.M1 := 0.0;
stGameTargetTorque.M2 := 0.0;
stGameTargetTorque.M3 := 0.0;


CASE eActiveGame OF

    E_GameID.PEELING:

        stGameTargetTorque :=
            fbPeelingGame.stJointTargetTorque;


    E_GameID.SORTER:

        stGameTargetTorque :=
            fbSorterGame.stJointTargetTorque;


    E_GameID.CRAZY_CAR:

        stGameTargetTorque :=
            fbCrazyCar.stJointTargetTorque;


    ELSE

        // No selected game generates torque

        stGameTargetTorque.M1 := 0.0;
        stGameTargetTorque.M2 := 0.0;
        stGameTargetTorque.M3 := 0.0;

END_CASE;

 




(*
		fbKinematic(q1:=GVL_RobotData.Q1_Actual, 
				q2:=GVL_RobotData.Q2_Actual,
				q3:=GVL_RobotData.Q3_Actual,
				X_Dir => xDir, 
				Y_Dir => yDir,
				Theta => theta,
				Beta => betaAngle);
				*)
				
	//eMode := E_RehabMode.Passive;
	
		 // Changing Operational Mode	
       // DoTaskSpaceControl();
	   
	   (*
	   
	   30 : (* ActiveMode *)
	   // Changing Operation mode  to CSV
	  IF bExecuteChangingMode THEN
			OperationalMode := En_TargetMode.eCSV;
   			fbSwitchMode(TargetMode := OperationalMode, Done => bSwitchopModeDone );
		END_IF
		
		IF  NOT bSwitchopModeDone  THEN
			
			bExecuteChangingMode := TRUE;
		ELSE
			bExecuteChangingMode := FALSE ; 
			eState :=34;
		END_IF

	34: // NEW STATE: CLEAR NC ERRORS
    fbMC_Reset1(Axis := GVL_Axes.Axis1, Execute := TRUE);
    fbMC_Reset2(Axis := GVL_Axes.Axis2, Execute := TRUE);
    fbMC_Reset3(Axis := GVL_Axes.Axis3, Execute := TRUE);

    IF fbMC_Reset1.Done AND fbMC_Reset2.Done AND fbMC_Reset3.Done THEN
        fbMC_Reset1(Axis := GVL_Axes.Axis1, Execute := FALSE);
        fbMC_Reset2(Axis := GVL_Axes.Axis2, Execute := FALSE);
		fbMC_Reset3(Axis := GVL_Axes.Axis3, Execute := FALSE);
        estate := 35; // Move to Enable only after NC is clear
    END_IF
		35: 
	fbMC_Power1.Enable := TRUE;
	fbMC_Power2.Enable := TRUE;    
	fbMC_Power3.Enable := TRUE;
    IF fbMC_Power1.Status AND fbMC_Power2.Status AND fbMC_Power3.Status THEN
        
        fbRobotisActive(bActiveModeIsDone => BActiveMode)  ;   // Now it is safe to execute the Jacobian control
    END_IF
	IF BActiveMode THEN
		eState := 40;
	END_IF
    
    // Safety check: if an error occurs, drop back to Passive
    IF RobotIsNotSafe THEN
        eState := 20;
	END_IF
	
	

		
    
    50: (* PREPARE FOR IMPEDANCE - Switch to CST *)
       

    60: (* RUN IMPEDANCE CONTROL *)
        // Note: In CST mode, you are sending raw torque commands to the drives
      IF fbMC_Power1.Status AND fbMC_Power2.Status AND fbMC_Power3.Status THEN
		  
		 fbRobotIsInIpedenceMode( bDone => ANNModeIsDone);
		 
	  END_IF

    IF ANNModeIsDone THEN
		eState := 70;
	END_IF
	
	*)
 
	 E_MainState.Fault: // motors disable
	 
	fbMC_Power1.Enable := FALSE;
	fbMC_Power2.Enable := FALSE;    
	fbMC_Power3.Enable := FALSE;
	   
END_CASE

END_PROGRAM

// ---- POUs/FB_DoHoming.TcPOU
FUNCTION_BLOCK FB_DoHoming
VAR_INPUT
	 HStart : BOOL;            (* Start homing *)
END_VAR
VAR_OUTPUT
	 HM123Done: BOOL;            (* Homing finished *)
	 HomingError : BOOL;
END_VAR
VAR
	 StateM1Homing : INT := 0;
	 StateM2M3Homing : INT := 0;
	 
   
   

    (* Velocity control FBs *)
    fbVelM1  : MC_MoveVelocity;
	fbVelM2  : MC_MoveVelocity;
    fbVelM3  : MC_MoveVelocity;
	fbMoReM1  : MC_MoveRelative;
	fbMoReM2  : MC_MoveRelative;
	fbMoReM3  : MC_MoveRelative;
	fbStopM1 : MC_Halt;
    fbStopM2 : MC_Halt;
    fbStopM3 : MC_Halt;
	
	

    (* Parameters *)
   	vBetaHome: LREAL:= 0.5; 			  (* safe speed for beta homing *)
	vThetaHome : LREAL := 0.5;    (* safe speed for theta homing *)
    vRHome     : LREAL := 0.5;    (* safe speed for R homing *)
	SwTheta1 : BOOL;
	SwR1: BOOL;
	
	
	StateM1: INT;
	SwBeta1: BOOL;
	HM1Done: BOOL;
	
	SwTheta2: BOOL;
	SwR2: BOOL;
	SwBeta2: BOOL;
	
	// Torque
	
    TorqueM1 : LREAL;
    TorqueM2 : LREAL;
    TorqueM3 : LREAL;
	TorqueLimitHome : LREAL := 60.0;
	tOverTorque : TON;
	fbStopLockM1: MC_STOP;
	fbStopLockM2: MC_STOP;
	fbStopLockM3: MC_STOP;
	
	// moves after contacting to Microswitch to reach nutral possition
	rSwBeta1  : R_TRIG;
	rSwTheta1 : R_TRIG;
	rSwR2 : R_TRIG;
	fbReadPosM1 : MC_ReadActualPosition;
	fbReadPosM2 : MC_ReadActualPosition;
	fbReadPosM3 : MC_ReadActualPosition;
	MinPosBeta: LREAL;
	
	NeutralOffsetBeta: LREAL;
	NutPosBeta: LREAL;
	MinPositionThM2: LREAL;
	NeutralOffsetM2: LREAL;
	NeutralOffsetM3: LREAL;
	MinPositionThM3: LREAL;
	MinPoTheta: LREAL;
	NeutralOffsetM2M3Theta: LREAL;
	NutPosTheta: LREAL;
	MinPositionRM2: LREAL;
	MinPositionRM3: LREAL;
	MinPoR: LREAL;
	NeutralOffsetM2M3R: LREAL;
	NutPosR: LREAL;
END_VAR


(* ========================== *)
(*       HOMING LOGIC         *)
(* ========================== *)

(* update switch values from global DWORD *)
SwTheta1 	 := (GVL_MicroSwitch.dwMicroSwitchDriverA AND 16#00020000) <> 0;  (* bit 0 *)
SwTheta2     := (GVL_MicroSwitch.dwMicroSwitchDriverA AND 16#00010000) <> 0;  (* bit 1 *)
SwR1    	 := (GVL_MicroSwitch.dwMicroSwitchDriverB AND 16#00080000) <> 0;  (* bit 0 *)
SwR2  		 := (GVL_MicroSwitch.dwMicroSwitchDriverB AND 16#00040000) <> 0;  (* bit 1 *)
SwBeta1      := (GVL_MicroSwitch.dwMicroSwitchDriverB AND 16#00020000) <> 0;  (* bit 2 *)
SwBeta2      := (GVL_MicroSwitch.dwMicroSwitchDriverB AND 16#00010000) <> 0;  (* bit 3 *)
		
			fbVelM1(
            Axis        := GVL_Axes.Axis1,
			velocity := vBetaHome,
			Acceleration := 1.0,
            Deceleration := 1000.0 );
			
			fbVelM2(
            Axis        := GVL_Axes.Axis2,
			velocity := vThetaHome,
			Acceleration := 1.0,
            Deceleration := 1000.0 );

        	fbVelM3(
            Axis        := GVL_Axes.Axis3,
			velocity := vThetaHome,
			Acceleration := 1.0,
            Deceleration := 1000.0 );
			
		fbStopM1(
            Axis         := GVL_Axes.Axis1,
            Deceleration := 1000.0);
		fbStopM2(
            Axis         := GVL_Axes.Axis2,
            Deceleration := 1000.0);
			
		fbStopM3(
            Axis         := GVL_Axes.Axis3,
            Deceleration := 1000.0);
			
		fbStopLockM1(
            Axis         := GVL_Axes.Axis1);
		fbStopLockM2(
            Axis         := GVL_Axes.Axis2);
		fbStopLockM3(
            Axis         := GVL_Axes.Axis3);	
			
			
// Reading Torque
TorqueM1 := GVL_Torque.TorqueM1_Act;
TorqueM2 := GVL_Torque.TorqueM2_Act;
TorqueM3 := GVL_Torque.TorqueM3_Act;	

// Reading Actual Position
fbReadPosM1(Axis := GVL_Axes.Axis1, Enable := TRUE);
fbReadPosM2(Axis := GVL_Axes.Axis2, Enable := TRUE);
fbReadPosM3(Axis := GVL_Axes.Axis3, Enable := TRUE);


// Mechanical Stopper
tOverTorque(
    IN := ABS(TorqueM1)  > TorqueLimitHome OR (ABS(TorqueM2)+ ABS(TorqueM3))  > TorqueLimitHome,
    PT := T#50MS);	
	IF toverTorque.Q  THEN
    (* stop all motors safely *)
    fbVelM1.Execute := FALSE;
    fbVelM2.Execute := FALSE;
    fbVelM3.Execute := FALSE;

    fbStopLockM1.Execute := TRUE;
    fbStopLockM2.Execute := TRUE;
	fbStopLockM3.Execute := TRUE;

    HomingError := TRUE;
       
END_IF

// Function Block - Move to Neutral Position
fbMoReM1(
 Axis:= GVL_Axes.Axis1,
 Velocity := vBetaHome,
 Acceleration := 10,
 Deceleration := 1000);
 
 fbMoReM2(
 Axis:= GVL_Axes.Axis2,
  Velocity := vThetaHome,
 Acceleration := 10,
 Deceleration := 1000);
 
 fbMoReM3(
 Axis:= GVL_Axes.Axis3,
 Velocity := vThetaHome,
 Acceleration := 10,
 Deceleration := 1000);
 
 

// Homing Motor A - Motor1
IF NOT HomingError THEN 
	
CASE StateM1Homing OF

    0:  (* IDLE *)
        HM1Done := FALSE;
        IF HStart THEN
            StateM1Homing := 10;      (* start beta homing *)
        END_IF


    10: (* HOME Beta: move pure -beta until SwBeta *)
        fbVelM1.Execute := TRUE;
		fbVelM1.Direction := MC_Direction.MC_Negative_Direction;
		rSwBeta1(CLK := SwBeta1);

         IF rSwBeta1.Q THEN 
                     
            MinPosBeta := fbReadPosM1.Position; 
		   	StateM1Homing := 15;
			
         
        END_IF
	
		
	15: (* WAIT UNTIL STOP AFTER THETA *)
        fbVelM1.Execute := FALSE;
		fbStopM1.Execute   := TRUE;
                 

        IF fbStopM1.Done THEN
            
            StateM1Homing := 17;   (* now ready for R homing *)
			NeutralOffsetBeta := ((121297.0/10000.0)/2) + ABS(fbReadPosM1.Position - MinPosBeta);
			
        END_IF
		
	17: (*Motor MOVE TO nutral position*)
	fbStopM1.Execute := FALSE;
    fbMoReM1.Execute := TRUE;
	fbMoReM1.Distance := NeutralOffsetBeta;
	
	IF fbMoReM1.Done THEN
		StateM1Homing := 20;
		NutPosBeta := fbReadPosM1.Position; 
		GVL_HomingResult.gHoming.HomePos_Beta :=NutPosBeta; 
	END_IF
	
	


    20: (* Homming of M1 is DONE *)
			
			fbMoReM1.Execute := FALSE;
			HM1Done := TRUE;

       
END_CASE





// Homing Motor B & C - (Motor 2 & 3)

CASE StateM2M3Homing OF

    0:  (* IDLE *)
        HM123Done := FALSE;

        IF HM1Done THEN
            StateM2M3Homing := 10;      (* start θ homing *)
        END_IF


    10: (* HOME THETA: move pure -theta until SwTheta *)
        fbVelM2.Execute := TRUE;
		fbVelM2.Direction := MC_Direction.MC_Positive_Direction;
		fbVelM3.Execute := TRUE;
		fbVelM3.Direction := MC_Direction.MC_Positive_Direction;
		rSwTheta1(CLK := SwTheta1);
		
		IF rSwTheta1.Q THEN 
                     
            MinPositionThM2 := fbReadPosM2.Position; 
			MinPositionThM3 := fbReadPosM3.Position;
			MinPoTheta := MinPositionThM2+MinPositionThM3;
		   	StateM2M3Homing := 15;
			
         
        END_IF
        
		
	15: (* WAIT UNTIL STOP AFTER THETA *)
			fbVelM2.Execute := FALSE;
			fbVelM3.Execute := FALSE;       
			fbStopM2.Execute   := TRUE;
      		fbStopM3.Execute   := TRUE;
            

        IF fbStopM2.Done AND fbStopM3.Done THEN
            
            StateM2M3Homing := 17;   (* now ready for R homing *)
			NeutralOffsetM2M3Theta := ((1.6384/360.0)*60.0) + MIN (ABS(fbReadPosM2.Position - MinPositionThM2), ABS(fbReadPosM3.Position - MinPositionThM3));
       // ((5000/10000)/2)
 END_IF
		
	17: (*Motors MOVE TO nutral position of THETA*)
		fbStopM2.Execute := FALSE;
		fbStopM3.Execute := FALSE;
		fbMoReM2.Execute := TRUE;
		fbMoReM3.Execute := TRUE;
		fbMoReM2.Distance := - NeutralOffsetM2M3Theta;
		fbMoReM3.Distance := - NeutralOffsetM2M3Theta;
		
	
	IF (fbMoReM2.Done AND fbMoReM3.Done) THEN
		StateM2M3Homing := 20;
		NutPosTheta := fbReadPosM2.Position + fbReadPosM3.Position; 
		GVL_HomingResult.gHoming.HomePos_Theta := NutPosTheta; 
	END_IF


    20: (* HOME R: move pure -R until SwR *)
		fbMoReM2.Execute := FALSE;
		fbMoReM3.Execute := FALSE; 
        fbVelM2.Execute   := TRUE;
		fbVelM2.Direction := MC_Direction.MC_Negative_Direction;
        fbVelM3.Execute   := TRUE;
		fbVelM3.Direction := MC_Direction.MC_Positive_Direction;
	
        rSwR2(CLK := SwR2);
		
		IF rSwR2.Q THEN 
                     
            MinPositionRM2 := fbReadPosM2.Position; 
			MinPositionRM3 := fbReadPosM3.Position;
			MinPoR := MinPositionRM2-MinPositionRM3;
			StateM2M3Homing := 25;
			
         END_IF
		 
	 
       

 
		
	25: (* WAIT UNTIL STOP AFTER R *)
		fbVelM3.Execute   := FALSE;
		fbVelM3.Execute   := FALSE;
        fbStopM2.Execute := TRUE;
        fbStopM3.Execute := TRUE;

        IF fbStopM2.Done AND fbStopM3.Done THEN
			
            
            StateM2M3Homing := 27;     (* finished homing *)
			NeutralOffsetM2M3R := (((16384.0/10000.0)/80.0)*5.0) + MIN (ABS(fbReadPosM2.Position - MinPositionRM2), ABS(fbReadPosM3.Position - MinPositionRM3));
        END_IF
		
	27: (*Motors MOVE TO nutral position of R*)
		fbStopM2.Execute := FALSE;
		fbStopM3.Execute := FALSE;
		fbMoReM2.Execute := TRUE;
		fbMoReM3.Execute := TRUE;
		fbMoReM2.Distance := NeutralOffsetM2M3R;
		fbMoReM3.Distance := -NeutralOffsetM2M3R;  // negative?
		
		IF (fbMoReM2.Done AND fbMoReM3.Done) THEN
		StateM2M3Homing := 30;
		NutPosR := fbReadPosM2.Position - fbReadPosM3.Position;
		GVL_HomingResult.gHoming.HomePos_R := NutPosR;  
	END_IF
	


    30: (* DONE *)
			fbMoReM2.Execute := FALSE;
			fbMoReM3.Execute := FALSE;
			fbStopM2.Execute   := FALSE;
        	fbStopM3.Execute   := FALSE;
       		HM123Done := TRUE;

        (* Wait for next cycle of HStart=FALSE before resetting *)
        IF NOT HStart THEN
            StateM2M3Homing := 0;   (* ready for next command *)
        END_IF

END_CASE

END_IF

END_FUNCTION_BLOCK

// ---- POUs/FB_ThreeAxisSafety.TcPOU
FUNCTION_BLOCK FB_ThreeAxisSafety
VAR_INPUT
	rDir : LREAL ;
	beta : LREAL ;
	theta : LREAL ;
		
END_VAR
VAR_OUTPUT
	AnyError   : BOOL;    (* live indication: some axis in error *)
END_VAR
  
VAR
	(* Status readbacks *)
    fbStatM1 : MC_ReadStatus;
    fbStatM2 : MC_ReadStatus;
    fbStatM3 : MC_ReadStatus;
	
	

    fbStopM1Safety : MC_Stop;
    fbStopM2Safety : MC_Stop;
    fbStopM3Safety : MC_Stop;
	

    anyErrInternal : BOOL;
	anyMicroswitchTrue: BOOL;
	//Errortype: STRING;
	// fbKinematicForSafety :FB_Kinematic;
	
END_VAR


(*
fbStopM1Safety(
            Axis         := GVL_Axes.Axis1,
			
            Deceleration := 1000.0);
		fbStopM2Safety(
            Axis         := GVL_Axes.Axis2,
            Deceleration := 1000.0);
			
		fbStopM3Safety(
            Axis         := GVL_Axes.Axis3,
            Deceleration := 1000.0);
fbKinematicForSafety(
    q1 := GVL_RobotData.Q1_Actual, 
    q2 := GVL_RobotData.Q2_Actual, 
    q3 := GVL_RobotData.Q3_Actual, 
 
    Theta => theta,
    R_Dir => rDir,
	Beta => beta    
);


(* === Read status of all three axes === *)
fbStatM1(
    Axis   := GVL_Axes.Axis1,
    Enable := TRUE);

fbStatM2(
    Axis   := GVL_Axes.Axis2,
    Enable := TRUE);

fbStatM3(
    Axis   := GVL_Axes.Axis3,
    Enable := TRUE);
	
// Micro_Switch
IF (GVL_MicroSwitch.dwMicroSwitchDriverA <> 0) OR (GVL_MicroSwitch.dwMicroSwitchDriverB <> 0) THEN
anyMicroswitchTrue := TRUE;
GVL_MessageStaus.MessageStaus := 'Microswitch is ON, Out OF ROM';
fbStopM1Safety.Execute :=TRUE;
		fbStopM2Safety.Execute :=TRUE;
		fbStopM3Safety.Execute :=TRUE;
		
END_IF

// OUT OF ROM
IF (rDir < 90 OR rDir > 468) OR 
   (beta < -60 OR beta > 60) OR 
   (theta < -30 OR theta > 30) THEN 
	 
GVL_MessageStaus.MessageStaus := 'OUT OF ROM';
		fbStopM1Safety.Execute :=TRUE;
		fbStopM2Safety.Execute :=TRUE;
		fbStopM3Safety.Execute :=TRUE;
END_IF
(* An axis is considered “in error” if ErrorStop is TRUE *)
anyErrInternal :=
       fbStatM1.Error
    OR fbStatM2.Error
    OR fbStatM3.Error
	OR (GVL_Axes.Axis1.NcToPlc.ErrorCode <> 0)
    OR (GVL_Axes.Axis2.NcToPlc.ErrorCode <> 0) 
    OR (GVL_Axes.Axis3.NcToPlc.ErrorCode <> 0);

(* === Stop command to all axes  === *)

IF anyErrInternal THEN

		
	GVL_MessageStaus.MessageStaus := 'Cycle Time Error';

END_IF

*)

END_FUNCTION_BLOCK

// ---- POUs/StopAllMotion.TcPOU
FUNCTION_BLOCK StopAllMotion
VAR_INPUT
	
END_VAR
VAR_OUTPUT
END_VAR

VAR
	MotionState : INT;
	fbStopM1 : MC_Stop;
    fbStopM2 : MC_Stop;
    fbStopM3 : MC_Stop;
	fbHaltM1 : MC_Halt;
	fbHaltM2 : MC_Halt;
	fbHaltM3 : MC_Halt;
END_VAR

IF GVL_HMI.EmergencyStopIsOnHardware THEN
	MotionState := 10;  // Pressed Hardware Emergency Stop
	
ELSIF GVL_HMI.EmergencyStopIsOnSoftware THEN
	MotionState := 20;	// Pressed software Emergency Stop
	
ELSE
	MotionState := 30;	// Deactivation All STOPS
	
END_IF



CASE MotionState OF

10:	

    fbStopM1(
        Axis      := GVL_Axes.Axis1,
        Execute   := TRUE);   

    fbStopM2(
        Axis      := GVL_Axes.Axis2,
        Execute   := TRUE);

    fbStopM3(
        Axis      := GVL_Axes.Axis3,
        Execute   := TRUE);
	
20:	
    fbHaltM1(
        Axis      := GVL_Axes.Axis1,
        Execute   := TRUE);   

    fbHaltM2(
        Axis      := GVL_Axes.Axis2,
        Execute   := TRUE);

    fbHaltM3(
        Axis      := GVL_Axes.Axis3,
        Execute   := TRUE);
30: 

 fbStopM1(
        Axis      := GVL_Axes.Axis1,
        Execute   := FALSE);   

    fbStopM2(
        Axis      := GVL_Axes.Axis2,
        Execute   := FALSE);

    fbStopM3(
        Axis      := GVL_Axes.Axis3,
        Execute   := FALSE);


 fbHaltM1(
        Axis      := GVL_Axes.Axis1,
        Execute   := FALSE);   

    fbHaltM2(
        Axis      := GVL_Axes.Axis2,
        Execute   := FALSE);

    fbHaltM3(
        Axis      := GVL_Axes.Axis3,
        Execute   := FALSE);

	
END_CASE

END_FUNCTION_BLOCK

// ---- POUs/FB_JointStateReader.TcPOU
FUNCTION_BLOCK FB_JointStateReader
VAR_INPUT
    Enable : BOOL := TRUE;
END_VAR

VAR_IN_OUT
    Axis1 : AXIS_REF;
    Axis2 : AXIS_REF;
    Axis3 : AXIS_REF;
END_VAR

VAR_OUTPUT
    JointState : ST_JointState; // Contains Position, Velocity, and Torque
END_VAR

VAR
    
END_VAR

// --- 1. Position (q1, q2, q3) ---
JointState.Position.q1     := Axis1.NcToPlc.ActPos;
JointState.Position.q2     := Axis2.NcToPlc.ActPos;
JointState.Position.q3     := Axis3.NcToPlc.ActPos;

// --- 2. Velocity (q1_dot, q2_dot, q3_dot) ---
JointState.Velocity.q1_dot := Axis1.NcToPlc.ActVelo;
JointState.Velocity.q2_dot := Axis2.NcToPlc.ActVelo;
JointState.Velocity.q3_dot := Axis3.NcToPlc.ActVelo;

// --- 3. Torque / Moment (M1, M2, M3) ---
JointState.Torque.M1       := Axis1.NcToPlc.ActTorque;
JointState.Torque.M2       := Axis2.NcToPlc.ActTorque;
JointState.Torque.M3       := Axis3.NcToPlc.ActTorque;

END_FUNCTION_BLOCK

// ---- POUs/FB_RobotKinematics.TcPOU
FUNCTION_BLOCK FB_RobotKinematics
VAR_INPUT
	JointData_INPUT : ST_JointState;
	CartesianData_INPUT : ST_CartesianState ;

END_VAR
VAR_OUTPUT
	JointData_Transed : ST_JointState;
	CartesianData_Transed : ST_CartesianState;
	Cartesian_PERCENTAGE_PoseObtainedFromForwardKinematic: ST_CartesianPose ;
	AdditionalPOSE : ST_CartesianAdditionalParametes;
END_VAR
VAR
	//JointPose : ST_JointPose;
//	ActBeta : LREAL;
	
//	ActR: LREAL;
 // Jacobian matrix
    J11 : LREAL;
    J12 : LREAL;
    J13 : LREAL;

    J21 : LREAL;
    J22 : LREAL;
    J23 : LREAL;

    J31 : LREAL;
    J32 : LREAL;
    J33 : LREAL;

	 
	
END_VAR


ForwardKinematics();


CalculateJacobian();

METHOD PUBLIC CalculateJacobian 
VAR_INPUT
//	 ActBeta : LREAL;
//	 ActR : LREAL;
	// JointVelo : ST_JointVelocity;
END_VAR

VAR
    // Local Variables
    BetaRad : LREAL;
    R_mm    : LREAL;
    PI_180    : LREAL := 0.0174532925199433; 
    

END_VAR
VAR_OUTPUT
	
	
	//CartesianVelocity : ST_CartesianVelocity;
	
	
	
END_VAR
BetaRad := AdditionalPOSE.BetaIncremental * PI_180; // Convert Degree to Radian
R_mm    := AdditionalPOSE.RIncremental;



J11 := -R_mm * GVL_ConstantCoefficent.K1 * PI_180 * COS(BetaRad); 
J12 :=  GVL_ConstantCoefficent.K2 * SIN(BetaRad);
J13 := -GVL_ConstantCoefficent.K2 * SIN(BetaRad);

// Row 2: How Y changes with motors
J21 :=  R_mm * GVL_ConstantCoefficent.K1 * PI_180 * SIN(BetaRad);
J22 :=  GVL_ConstantCoefficent.K2 * COS(BetaRad);
J23 := -GVL_ConstantCoefficent.K2 * COS(BetaRad);

// Row 3: How Theta (Wrist) changes with motors
J31 := 0.0;
J32 := -GVL_ConstantCoefficent.K3 / 2.0;
J33 := -GVL_ConstantCoefficent.K3 / 2.0;

CartesianData_Transed.Velocity.Vx := J11* JointData_INPUT.Velocity.q1_dot + J12* JointData_INPUT.Velocity.q2_dot + J13* JointData_INPUT.Velocity.q3_dot;
CartesianData_Transed.Velocity.Vy := J21* JointData_INPUT.Velocity.q1_dot + J22* JointData_INPUT.Velocity.q2_dot + J23* JointData_INPUT.Velocity.q3_dot;
CartesianData_Transed.Velocity.Vtheta := J31* JointData_INPUT.Velocity.q1_dot + J32* JointData_INPUT.Velocity.q2_dot + J33* JointData_INPUT.Velocity.q3_dot;


// JacobianTrans
//JointData_Transed.Torque.M1 := J11* CartesianData_INPUT.Force.Fx + J21* CartesianData_INPUT.Force.Fy+ J31* CartesianData_INPUT.Force.Mtheta;
//JointData_Transed.Torque.M2 := J12* CartesianData_INPUT.Force.Fx + J22* CartesianData_INPUT.Force.Fy+ J32* CartesianData_INPUT.Force.Mtheta;
//JointData_Transed.Torque.M3 := J13* CartesianData_INPUT.Force.Fx + J23* CartesianData_INPUT.Force.Fy+ J33* CartesianData_INPUT.Force.Mtheta;
END_METHOD

METHOD PUBLIC CartesianForceToTorque
VAR_INPUT
    Force : ST_CartesianForces;
END_VAR

VAR_OUTPUT
    Torque : ST_JointTorque;
END_VAR
Torque.M1 :=
      J11 * Force.Fx
    + J21 * Force.Fy
    + J31 * Force.Mtheta;

Torque.M2 :=
      J12 * Force.Fx
    + J22 * Force.Fy
    + J32 * Force.Mtheta;

Torque.M3 :=
      J13 * Force.Fx
    + J23 * Force.Fy
    + J33 * Force.Mtheta;
END_METHOD

METHOD PUBLIC ForwardKinematics : BOOL
VAR_INPUT
//	JointPose : ST_JointPose;
END_VAR

VAR
Theta : LREAL;
	R_Dir : LREAL;
	X_Dir : LREAL;	
	Y_Dir : LREAL;
	Beta : LREAL;
	X0: LREAL;
	Y0: LREAL;
	X1: LREAL;
	LineLength: INT := 5;
	Y1: LREAL;
	
	// Test Visualization
	A : INT := 1000;
	B : INT := 1000;
	C : INT;
	D: LREAL;
	E : LREAL;
	
	R_Visu: INT;
	Theta_Visu: INT;
	X_Visu: INT;
	Y_Visu: INT;
	X_Dir_Abs: LREAL;
	Y_Dir_Abs: LREAL;
	R_Dir_Abs: LREAL;
	WristAngle: LREAL;
	WristAngle_Abs: LREAL;
	
	BetaFromAbsolute : LREAL;
	ThetaFromAbsolute : LREAL;
	LinearFromAbsolute : LREAL;
	
	END_VAR
VAR_OUTPUT
	//CartesianPoseObtainedFromForwardKinematic : ST_CartesianPose;
	//	Cartesian_PERCENTAGE_PoseObtainedFromForwardKinematic: ST_CartesianPose ; 
	//CartesianAdditionalPose: ST_CartesianAdditionalParametes ;
END_VAR

// Forward Kinematic From Incremental Encoders

R_Dir := 464.0 -  GVL_ConstantCoefficent.K2*(JointData_INPUT.Position.q2-JointData_INPUT.Position.q3-GVL_HomingResult.gHoming.HomePos_R);   // Unit : mm 
Theta := -GVL_ConstantCoefficent.K3*(JointData_INPUT.Position.q2+JointData_INPUT.Position.q3-GVL_HomingResult.gHoming.HomePos_Theta)/2.0; // Unid: Degree
Beta := GVL_ConstantCoefficent.K1*(JointData_INPUT.Position.q1-GVL_HomingResult.gHoming.HomePos_Beta);

X_Dir := R_Dir * (SIN(- Beta * (PI / 180.0)));   // 464 is maximum R
Y_Dir := 464 -(R_Dir  * (COS(Beta * (PI / 180.0))));
Y_Dir := 464.0 -(R_Dir  * (COS(Beta * (PI / 180.0))));
WristAngle := Theta;

CartesianData_Transed.Position.X := X_Dir;
CartesianData_Transed.Position.Y := Y_Dir;
CartesianData_Transed.Position.Theta := WristAngle;

// NORMALIZATION OF INCREMENTAL DATA
// 1. Normalize Y_Dir (0-370mm) to Percentage (0-100)
// We check for negative values just in case calibration is slightly off
IF Y_Dir < 0.0 THEN 
    Cartesian_PERCENTAGE_PoseObtainedFromForwardKinematic.Y := 0.0;
ELSIF Y_Dir > 370.0 THEN 
    Cartesian_PERCENTAGE_PoseObtainedFromForwardKinematic.Y := 100.0;
ELSE
    // The main formula: (Current / Max) * 100
    Cartesian_PERCENTAGE_PoseObtainedFromForwardKinematic.Y := (Y_Dir / 370.0) * 100.0;
END_IF

IF X_Dir < -410.0 THEN 
    Cartesian_PERCENTAGE_PoseObtainedFromForwardKinematic.X := -100.0;
ELSIF X_Dir > 410.0 THEN 
    Cartesian_PERCENTAGE_PoseObtainedFromForwardKinematic.X := 100.0;
ELSE
    // The main formula: (Current / Max) * 100
    Cartesian_PERCENTAGE_PoseObtainedFromForwardKinematic.X := (X_Dir / 410.0) * 100.0;
END_IF


(*
GVL_EndeffectorPosition.R_Dir := 464.0 -  GVL_ConstantCoefficent.K2*(JointPose.q2-JointPose.q3-GVL_HomingResult.gHoming.HomePos_R);   // Unit : mm 
Theta := -GVL_ConstantCoefficent.K3*(JointPose.q2+JointPose.q3-GVL_HomingResult.gHoming.HomePos_Theta)/2.0; // Unid: Degree
CartesianAdditionalPose.BetaIncremental := GVL_ConstantCoefficent.K1*(JointPose.q1-GVL_HomingResult.gHoming.HomePos_Beta);

CartesianPose.X := R_Dir * (SIN(- Beta * (PI / 180.0)));   // 464 is maximum R
CartesianPose.Y := 464.0 -(R_Dir  * (COS(Beta * (PI / 180.0))));
CartesianPose.Theta := Theta;

*)

// Absolute Encoder




BetaFromAbsolute :=  (TO_LREAL(GVL_AbsoluteEncoders.AbsoluteBetaPosition) / 16384.0) * 360.0;
LinearFromAbsolute :=  (TO_LREAL(GVL_AbsoluteEncoders.AbsoluteLinearPosition) / 4096.0);  //mm
ThetaFromAbsolute :=  (TO_LREAL(GVL_AbsoluteEncoders.AbsoluteTetaPosition) / 16384.0) * 360.0;  // This is wrist Angle
R_Dir_Abs := 464.0 -(LinearFromAbsolute + 402.7); // 464 comes from solidworks , 402.7 comes from absoute encodere date when robot placed in home position, if there is a about1-2 mm error between what i read from incremental and absolute can have a roote here, but this error should be constant, if during motion the numbers changed is related your code or shows slipping of cable!

AdditionalPOSE.X_Dir_Abs := R_Dir_Abs * (SIN((-BetaFromAbsolute - 114.16) * (PI / 180.0)));   // 464 is maximum R, 114.16 is shifting number I read whem robot placed in home position 
AdditionalPOSE.Y_Dir_Abs := 464.0 -(R_Dir_Abs  * (COS((-BetaFromAbsolute - 114.16) * (PI / 180.0))));
AdditionalPOSE.WristAngle_Abs := ThetaFromAbsolute;
AdditionalPOSE.RIncremental := R_Dir ;
AdditionalPOSE.BetaIncremental := Beta;






(*   Between * hidden because it is related to games and visualization

//PONG GAME
// 1. Normalize Y_Dir (0-370mm) to Percentage (0-100)
// We check for negative values just in case calibration is slightly off
IF Y_Dir < 0 THEN 
    GVL_GamePong.MyRobotY := 0;
ELSIF Y_Dir > 370 THEN 
    GVL_GamePong.MyRobotY := 100;
ELSE
    // The main formula: (Current / Max) * 100
    GVL_GamePong.MyRobotY := TO_REAL((Y_Dir / 370.0) * 100.0);
END_IF




// Wrist Rotation visualization

Theta_Visu := TO_INT(Theta) + TO_INT(Beta);

// linear of visualizartion
*)

//E :=  - (R_Dir*10);
//R_Visu := TO_INT(E);
GVL_HMI.EndeffectorPositionPixcelUnit_X := TO_INT(CartesianData_Transed.Position.X * (245.0/375.0))+500-7;
GVL_HMI.EndeffectorPositionPixcelUnit_Y := -TO_INT(CartesianData_Transed.Position.Y * ((245.0/375.0)))+687-7;
GVL_HMI.EndeffectorPositionPixcelUnit_Theta := WristAngle;
END_METHOD

END_FUNCTION_BLOCK

// ---- POUs/FB_RobotIsActive.TcPOU
FUNCTION_BLOCK FB_RobotIsActive
VAR_INPUT
	


END_VAR
VAR_OUTPUT
	bBusy         : BOOL;
    bDone         : BOOL;
    // Final CSV commands to the drives
    lrTargetVelX  : LREAL; 
    lrTargetVelY  : LREAL;
    lrTargetVelTheta : LREAL;
	bActiveModeIsDone : BOOL;
END_VAR
VAR
	
(* Variables for UpdatePathPlanning *)
// Segment Lengths
    lrL1, lrL2, lrL3 : LREAL;
    
    // Direction Unit Vectors
    lrDX1, lrDY1, lrDTh1 : LREAL;
    lrDX2, lrDY2, lrDTh2 : LREAL;
    lrDX3, lrDY3, lrDTh3 : LREAL;
    
    // Feedforward Velocity Outputs
    lrVx_FF, lrVy_FF, lrVTh_FF : LREAL;
	
	iCurrentSegment : INT; // 10 for A-B, 20 for B-C, 30 for C-A
(*----------------------------------------*)



	
    stPointA      : ARRAY[1..3] OF LREAL := [100,100,0]; // [X, Y, Theta]
    stPointB      : ARRAY[1..3] OF LREAL := [-200,200,0];
    stPointC      : ARRAY[1..3] OF LREAL := [100,200,0];
    lrVmax        : LREAL := 10 ; // Max Velocity (mm/s)
    lrAcc         : LREAL := 20 ; // Symmetrical Acc/Dec (mm/s^2)
	
	// Feedback from Motors (mapped from EPOS4 PDOs)
	// fbKinematic : FB_Kinematic;
	
    lrActX        : LREAL ; 
    lrActY        : LREAL ;
    lrActTheta    : LREAL ;
 	lrActR    : LREAL ;



iState        : INT;    // State Machine index
    fbWaitTimer   : TON;    // 1-second pause timer
    lrS_T         : LREAL;  // Current path distance
    lrS_dot       : LREAL;  // Current path velocity (Feedforward)
    
    // Internal setpoints calculated each cycle
    stCurrentSet  : ARRAY[1..3] OF LREAL; // Target [X, Y, Theta]
    
  
   
	(*PID Controller Using Tc2_ControllerToolbox*)
	
	// PID Instances
    fbPidX, fbPidY, fbPidTheta : FB_CTRL_PID;
    
    // Parameter Structures (Required for FB_CTRL_PID)
    stParamsX, stParamsY, stParamsTheta : ST_CTRL_PID_PARAMS;
    
    // The mode variable to turn them on/off
    eMode : E_CTRL_MODE;
	
	
	// Final Control Outputs (Sent to Jacobian/Motors)
    lrVx_Total    : LREAL;
    lrVy_Total    : LREAL;
    lrVTh_Total   : LREAL;

	
	(*-----------------------------------*)
	
	// Final joint targets to be sent to motors
    JointVelTarget : ARRAY[1..3] OF LREAL;
	
	
	
	
	// Triangle Path
	
	State : INT;
	X_S: LREAL;
	S_T: LREAL; // Current position setpoint
	dx: LREAL;
	dy: LREAL;
	L: LREAL;
	Y_S: LREAL;
	dx1: LREAL;
	dy1: LREAL;
	L1: LREAL;
	dx2: LREAL;
	dy2: LREAL;
	L2: LREAL;
	dx3: LREAL;
	dy3: LREAL;
	L3: LREAL;
	dTh1: LREAL;
	dTh2: LREAL;
	dTh3: LREAL;
	Theta_S: LREAL;
	
	// S(t) definition
	 
    S_dot    : LREAL; // Current velocity (Feedforward)
	lrL_Target: LREAL;
	bSegmentDone: BOOL;
	//MessageStaus : STRING(255); 
	
	bAtPointA: BOOL;
	lrApproachStartX: LREAL;
	lrApproachStartY: LREAL;
	lrApproachStartTheta: LREAL;
	lrDX_App: LREAL;
	lrDY_App: LREAL;
	lrDTh_App: LREAL;
	lrL_App: LREAL;
	bWaitEnable: BOOL := FALSE;
END_VAR

(*
fbKinematic(
    q1 := GVL_RobotData.Q1_Actual, 
    q2 := GVL_RobotData.Q2_Actual, 
    q3 := GVL_RobotData.Q3_Actual, 
    X_Dir => lrActX, 
    Y_Dir => lrActY, 
    Theta => lrActTheta,
	R_Dir => lrActR    
);

fbWaitTimer(
    IN := bWaitEnable,
    PT := T#50S
);
CASE iState OF
	0: // Initialization State
        
            
// Initialization for Approchig to A point 

// 1. Capture the exact starting position of the robot right now
lrApproachStartX     := lrActX;
lrApproachStartY     := lrActY;
lrApproachStartTheta := lrActTheta;

// 2. Calculate the distance and direction to Point A
lrDX_App  := stPointA[1] - lrApproachStartX;
lrDY_App  := stPointA[2] - lrApproachStartY;
lrDTh_App := stPointA[3] - lrApproachStartTheta;

// 3. Calculate the total approach length
lrL_App   := MAX(0.001, SQRT(lrDX_App*lrDX_App + lrDY_App*lrDY_App));

// 4. Update the status message for the GUI


// --- Line 1: A to B ---
            lrDX1  := stPointB[1] - stPointA[1];
            lrDY1  := stPointB[2] - stPointA[2];
            lrDTh1 := stPointB[3] - stPointA[3];
            lrL1   := MAX(0.001, SQRT(lrDX1*lrDX1 + lrDY1*lrDY1));
            
            // --- Line 2: B to C ---
            lrDX2  := stPointC[1] - stPointB[1];
            lrDY2  := stPointC[2] - stPointB[2];
            lrDTh2 := stPointC[3] - stPointB[3];
            lrL2   := MAX(0.001, SQRT(lrDX2*lrDX2 + lrDY2*lrDY2));
            
            // --- Line 3: C to A ---
            lrDX3  := stPointA[1] - stPointC[1];
            lrDY3  := stPointA[2] - stPointC[2];
            lrDTh3 := stPointA[3] - stPointC[3];
            lrL3   := MAX(0.001, SQRT(lrDX3*lrDX3 + lrDY3*lrDY3));
			
			
            
            // --- Reset Global Motion Variables ---
            lrS_T   := 0; // Current distance along path
            lrS_dot := 0; // Current velocity
			
			// PID SEction
			// 1. Setup X-Axis Parameters
        stParamsX.tCtrlCycleTime := T#10MS;
        stParamsX.tTaskCycleTime := T#10MS;
        stParamsX.fKp            := 1.5;   // Proportional Gain
        stParamsX.tTn            := T#100MS; // Integral Time
        stParamsX.fOutMaxLimit   := 100;   // Safety: Max speed limit (mm/s)
        stParamsX.fOutMinLimit   := -100;
        
        // 2. Setup Y and Theta (Using same parameters or unique ones)
        stParamsY     := stParamsX;
        stParamsTheta := stParamsX;
        
        // 3. Set the mode to Active for the controllers
        eMode := eCTRL_MODE_ACTIVE;
           iCurrentSegment := 5;
		   GVL_MessageStaus.MessageStaus := 'Robot is approaching Point A.';
            iState  := 5; // Approching to A point 
        
		
	
5: // --- APPROACH: Move to Point A ---
    // Stage 1: Trajectory
    bAtPointA := UpdateTrapezoid(lrL_total := lrL_App);

    // Stage 2: Path Mapping (Manual mapping for this one-time move)
    stCurrentSet[1] := lrApproachStartX + (lrDX_App / lrL_App) * lrS_T;
    stCurrentSet[2] := lrApproachStartY + (lrDY_App / lrL_App) * lrS_T;
    stCurrentSet[3] := lrApproachStartTheta + (lrDTh_App / lrL_App) * lrS_T;
    
    lrVx_FF := (lrDX_App / lrL_App) * lrS_dot;
    lrVy_FF := (lrDY_App / lrL_App) * lrS_dot;
    lrVTh_FF := (lrDTh_App / lrL_App) * lrS_dot;

    // Stages 3, 4, 5: ControlLoop, Jacobian, DriveMotors (Call as normal)
   ControlLoop();

    // STAGE 4: Solving Inverse Jacobian
    // Transforms Cartesian totals into joint velocities (dqTarget)
    IF CalculateInverseJacobian(
        TargetVelX     := lrVx_Total, 
        TargetVelY     := lrVy_Total, 
        TargetVelTheta := lrVTh_Total,
        ActR           := lrActR, 
        ActTheta       := lrActTheta
    ) THEN
        
        // STAGE 5: Drive Motors
        DriveMotors(bEnableMotion := TRUE);
		
	END_IF
	IF bAtPointA THEN
		GVL_MessageStaus.MessageStaus  := 'Robot is Reached A.';
		bWaitEnable := TRUE;   // start TON;
		
		iState := 7;
	END_IF



7: // Waiting before Start A-B movement

GVL_MessageStaus.MessageStaus  := 'Waiting For start Main active path';
  DriveMotors(bEnableMotion := FALSE);

    IF fbWaitTimer.Q THEN
       bWaitEnable := FALSE;
		lrS_T := 0;             // Reset progress for the triangle
        lrS_dot := 0;
        iCurrentSegment := 10;  // Set for Line A -> B
        iState := 10;           // Start the main task
		GVL_MessageStaus.MessageStaus  := 'Robot is Moving from  A To B.';
    END_IF

10:	
	// --- CONSOLIDATED ACTIVE MOTION (A -> B -> C -> A) ---

    // STAGE 1: Trajectory Planning
    // Use a target distance based on the current segment
    CASE iCurrentSegment OF
        10: lrL_Target := lrL1;
        20: lrL_Target := lrL2;
        30: lrL_Target := lrL3;
    END_CASE

    // Updates lrS_T and lrS_dot. Returns TRUE when target is reached.
    bSegmentDone := UpdateTrapezoid(lrL_total := lrL_Target);

    // STAGE 2: Path Mapping
    // Uses the iCurrentSegment to pick the right dX, dY, dTh and calculate FF
    UpdatePathSetpoints();

    // STAGE 3: Control Loop (PID)
    // Results in lrVx_Total, lrVy_Total, lrVTh_Total
    ControlLoop();

    // STAGE 4: Solving Inverse Jacobian
    // Transforms Cartesian totals into joint velocities (dqTarget)
    IF CalculateInverseJacobian(
        TargetVelX     := lrVx_Total, 
        TargetVelY     := lrVy_Total, 
        TargetVelTheta := lrVTh_Total,
        ActR           := lrActR, 
        ActTheta       := lrActTheta
    ) THEN
        
        // STAGE 5: Drive Motors
        DriveMotors(bEnableMotion := TRUE);
        
    END_IF

    // --- AUTOMATIC SEGMENT TRANSITION ---
 IF bSegmentDone THEN
    bWaitEnable := TRUE; 
	lrS_T       := 0;     // Safe to reset path distance
    lrS_dot     := 0;     // Safe to reset velocity ramp
END_IF

// 2. While the timer is active, override motion to 0.0
IF bWaitEnable THEN
    DriveMotors(bEnableMotion := FALSE); // Use your "Active Zero" logic
	

END_IF

// 3. Monitor the timer independently of the 'Done' flag
IF fbWaitTimer.Q THEN
    bWaitEnable := FALSE; // Reset timer for next corner
    
    
    // Increment Segment
    IF iCurrentSegment = 10 THEN
        iCurrentSegment := 20;
        GVL_MessageStaus.MessageStaus := 'Moving B to C.';
    ELSIF iCurrentSegment = 20 THEN
        iCurrentSegment := 30;
        GVL_MessageStaus.MessageStaus := 'Moving C to A.';
    ELSIF iCurrentSegment = 30 THEN
        iState := 40; // End of triangle
        GVL_MessageStaus.MessageStaus := 'Task finished.';
    END_IF
END_IF
	
	40: // Entire Triangle Complete
       bActiveModeIsDone := TRUE;
		
END_CASE
*)

METHOD CalculateInverseJacobian : BOOL
VAR_INPUT
    // Values passed from your State Machine or PID controllers
    TargetVelX     : LREAL; 
    TargetVelY     : LREAL; 
    TargetVelTheta : LREAL; 
	ActR           : LREAL; // Pass current R position here
    ActTheta       : LREAL; // Pass current Beta/Theta position here
END_VAR
VAR
    // Temporary variables used ONLY for this calculation
    BetaRad   : LREAL;
    R_mm      : LREAL;
    DotR      : LREAL; 
    PI_180    : LREAL := 0.0174532925199433; 
END_VAR
// 1. Assign local values from FB or GVL sources
BetaRad := ActTheta * PI_180;
R_mm    := ActR;

// 2. Singularity Protection
IF R_mm < 0.1 THEN
    JointVelTarget[1] := 0.0;
    JointVelTarget[2] := 0.0;
    JointVelTarget[3] := 0.0;
    CalculateInverseJacobian := FALSE;
    RETURN;
END_IF

// 3. Intermediate Radial Velocity
DotR := (TargetVelX * SIN(-BetaRad)) - (TargetVelY * COS(BetaRad));

// 4. Calculate Final Outputs (Stored in FB's JointVelTarget array)
JointVelTarget[1] := (-TargetVelX * COS(BetaRad) - TargetVelY * SIN(-BetaRad)) 
                      / (GVL_ConstantCoefficent.K1 * PI_180 * R_mm);

JointVelTarget[2] := (TargetVelTheta / -GVL_ConstantCoefficent.K3) + (DotR / (-2.0 * GVL_ConstantCoefficent.K2));
JointVelTarget[3] := (TargetVelTheta / -GVL_ConstantCoefficent.K3) - (DotR / (-2.0 * GVL_ConstantCoefficent.K2));

CalculateInverseJacobian := TRUE;
END_METHOD

METHOD ControlLoop : BOOL
// 1. AXIS X CONTROL
fbPidX(
    fSetpointValue := stCurrentSet[1], // From your Path Planning
    fActualValue   := lrActX,          // From Forward Kinematics
    eMode          := eMode,           // Defined in your VAR section
    stParams       := stParamsX        // Parameters from State 0
);
// Total Velocity = Feedforward + PID correction
lrVx_Total := lrVx_FF + fbPidX.fOut; 

// 2. AXIS Y CONTROL
fbPidY(
    fSetpointValue := stCurrentSet[2], 
    fActualValue   := lrActY, 
    eMode          := eMode, 
    stParams       := stParamsY
);
lrVy_Total := lrVy_FF + fbPidY.fOut;

// 3. AXIS THETA CONTROL
fbPidTheta(
    fSetpointValue := stCurrentSet[3], 
    fActualValue   := lrActTheta, 
    eMode          := eMode, 
    stParams       := stParamsTheta
);
lrVTh_Total := lrVTh_FF + fbPidTheta.fOut;




ControlLoop := TRUE;
END_METHOD

METHOD DriveMotors : BOOL
VAR_INPUT
	bEnableMotion : BOOL;
END_VAR
VAR
    fbMoveVel_Axis1 : MC_MoveVelocity;
    fbMoveVel_Axis2 : MC_MoveVelocity;
    fbMoveVel_Axis3 : MC_MoveVelocity;
	numM1Direction : MC_Direction;
	numM2Direction : MC_Direction;
	numM3Direction : MC_Direction;
	
	
	lrTargetVelM1: LREAL;
	lrTargetVelM2 : LREAL;
	lrTargetVelM3 : LREAL;
END_VAR
// 1. Determine Direction for Axis 1 based on Jacobian Output
IF JointVelTarget[1] >= 0 THEN
    numM1Direction := MC_Positive_Direction;
ELSE
    numM1Direction := MC_Negative_Direction;
END_IF

// 2. Execute Axis 1 Motion
IF bEnableMotion THEN
    lrTargetVelM1 := ABS(JointVelTarget[1]);
	
ELSE
    lrTargetVelM1 := 0.0; // Force zero during state 7
END_IF
fbMoveVel_Axis1(
    Axis          := GVL_Axes.Axis1,
    Execute       := TRUE, 
    Velocity      := lrTargetVelM1 ,   // Use Absolute value since direction is explicit
    Acceleration  := lrAcc,              // Acc/Dec must always be positive
    Deceleration  := lrAcc, 
    Direction     := numM1Direction,     // Explicitly set to Positive or Negative
    BufferMode    := MC_Aborting
);

// 3. Repeat Logic for Axis 2
IF JointVelTarget[2] >= 0 THEN
    numM2Direction := MC_Positive_Direction;
ELSE
    numM2Direction := MC_Negative_Direction;
END_IF

IF bEnableMotion THEN
    lrTargetVelM2 := ABS(JointVelTarget[2]);
	
ELSE
    lrTargetVelM2 := 0.0; // Force zero during state 7
END_IF

fbMoveVel_Axis2(
    Axis          := GVL_Axes.Axis2,
    Execute       := TRUE,
    Velocity      := lrTargetVelM2,
    Acceleration  := lrAcc,
    Deceleration  := lrAcc,
    Direction     := numM2Direction
);

// 4. Repeat Logic for Axis 3
IF JointVelTarget[3] >= 0 THEN
    numM3Direction := MC_Positive_Direction;
ELSE
    numM3Direction := MC_Negative_Direction;
END_IF
IF bEnableMotion THEN
    lrTargetVelM3 := ABS(JointVelTarget[3]);
	
ELSE
    lrTargetVelM3 := 0.0; // Force zero during state 7
END_IF
fbMoveVel_Axis3(
    Axis          := GVL_Axes.Axis3,
    Execute       := TRUE,
    Velocity      := lrTargetVelM3,
    Acceleration  := lrAcc,
    Deceleration  := lrAcc,
    Direction     := numM3Direction
);
END_METHOD

METHOD UpdatePathSetpoints : BOOL
VAR_INPUT
END_VAR

CASE iCurrentSegment OF
    10: // Line A -> B
        IF lrL1 > 0.0 THEN
            stCurrentSet[1] := stPointA[1] + (lrDX1 / lrL1) * lrS_T;
            stCurrentSet[2] := stPointA[2] + (lrDY1 / lrL1) * lrS_T;
            stCurrentSet[3] := stPointA[3] + (lrDTh1 / lrL1) * lrS_T;
            
            // Calculate Feedforward Velocities (Unit Vector * Current Speed)
            lrVx_FF := (lrDX1 / lrL1) * lrS_dot;
            lrVy_FF := (lrDY1 / lrL1) * lrS_dot;
            lrVTh_FF := (lrDTh1 / lrL1) * lrS_dot;
        END_IF;

    20: // Line B -> C
        IF lrL2 > 0.0 THEN
            stCurrentSet[1] := stPointB[1] + (lrDX2 / lrL2) * lrS_T;
            stCurrentSet[2] := stPointB[2] + (lrDY2 / lrL2) * lrS_T;
            stCurrentSet[3] := stPointB[3] + (lrDTh2 / lrL2) * lrS_T;
            
            lrVx_FF := (lrDX2 / lrL2) * lrS_dot;
            lrVy_FF := (lrDY2 / lrL2) * lrS_dot;
            lrVTh_FF := (lrDTh2 / lrL2) * lrS_dot;
        END_IF;

    30: // Line C -> A
        IF lrL3 > 0.0 THEN
            stCurrentSet[1] := stPointC[1] + (lrDX3 / lrL3) * lrS_T;
            stCurrentSet[2] := stPointC[2] + (lrDY3 / lrL3) * lrS_T;
            stCurrentSet[3] := stPointC[3] + (lrDTh3 / lrL3) * lrS_T;
            
            lrVx_FF := (lrDX3 / lrL3) * lrS_dot;
            lrVy_FF := (lrDY3 / lrL3) * lrS_dot;
            lrVTh_FF := (lrDTh3 / lrL3) * lrS_dot;
        END_IF;
END_CASE
END_METHOD

METHOD UpdateTrapezoid : BOOL
VAR_INPUT
	lrL_total : LREAL;
	
END_VAR

VAR
		
    dist_rem  : LREAL;
    CycleTime : LREAL := 0.01;  //plc cycle time is 10 ms
	S_dec : LREAL; // calcullated stopping distance
	
END_VAR
// This method calculates the current velocity and distance scalar for the move.

s_dec := (lrVmax * lrVmax) / (2.0 * lrAcc);
dist_rem := lrL_total - lrS_T;

IF dist_rem > s_dec THEN
    lrS_dot := MIN(lrS_dot + (lrAcc * CycleTime), lrVmax);
ELSE
    lrS_dot := SQRT(2.0 * lrAcc * MAX(0.0, dist_rem));
END_IF

lrS_T := lrS_T + (lrS_dot * CycleTime);

IF dist_rem <= 0.001 THEN
    UpdateTrapezoid := TRUE; // Signal segment complete
END_IF
END_METHOD

END_FUNCTION_BLOCK

// ---- POUs/FB_SwitchOpMode.TcPOU
FUNCTION_BLOCK FB_SwitchOpMode
VAR_INPUT
		
    TargetMode       : En_TargetMode;   // ENUM instead of magic numbers
   
END_VAR
VAR_OUTPUT
	Done  : BOOL;
    Busy  : BOOL;
    Error : BOOL;
	
END_VAR
VAR
	fbDisable : MC_Power;
    fbEnable  : MC_Power;
    state     : INT := 0;
	tWait    : TON;
	fbStopM1 : MC_Halt;
	fbStopM2 : MC_Halt;
	fbStopM3 : MC_Halt;
	fbPowerM1 : MC_Power ;
	fbPowerM2 : MC_Power ;
	fbPowerM3 : MC_Power ;
	fbWriteModeM1 : MC_WriteDriveOperationMode;
	fbWriteModeM2 : MC_WriteDriveOperationMode;
	fbWriteModeM3 : MC_WriteDriveOperationMode;
	DriveOperationMode : E_DriveOperationMode;
	
	fbReadModeM1 :  MC_ReadDriveOperationMode;
	fbReadModeM2 :  MC_ReadDriveOperationMode;
	fbReadModeM3 :  MC_ReadDriveOperationMode;
	
	
	bStopCmd: BOOL;
	bPowerEnable: BOOL;
	bWriteMode: BOOL;
	bWait: BOOL;
	bReadMode: BOOL;
	Test : ARRAY [1..5] OF INT; 
	Testii: INT := 1;
	LastErrorCode: UDINT;
END_VAR

	
	// ===== FB calls (always executed) =====

fbStopM1(Axis := GVL_Axes.Axis1, Execute := bStopCmd, Deceleration := 100.0);
fbStopM2(Axis := GVL_Axes.Axis2, Execute := bStopCmd, Deceleration := 100.0);
fbStopM3(Axis := GVL_Axes.Axis3, Execute := bStopCmd, Deceleration := 100.0);

fbPowerM1(Axis := GVL_Axes.Axis1, Enable := bPowerEnable);
fbPowerM2(Axis := GVL_Axes.Axis2, Enable := bPowerEnable);
fbPowerM3(Axis := GVL_Axes.Axis3, Enable := bPowerEnable);

fbWriteModeM1(
    Axis := GVL_Axes.Axis1,
    Execute := bWriteMode,
    DriveOperationMode := TO_SINT(TargetMode)
);
fbWriteModeM2(
    Axis := GVL_Axes.Axis2,
    Execute := bWriteMode,
    DriveOperationMode := TO_SINT(TargetMode)
);
fbWriteModeM3(
    Axis := GVL_Axes.Axis3,
    Execute := bWriteMode,
    DriveOperationMode := TO_SINT(TargetMode)
);

fbReadModeM1(
    Axis := GVL_Axes.Axis1,
    Execute := bReadMode
);

fbReadModeM2(
    Axis := GVL_Axes.Axis2,
    Execute := bReadMode
);

fbReadModeM3(
    Axis := GVL_Axes.Axis3,
    Execute := bReadMode
);



tWait(IN := bWait, PT := T#1S);
	
	
CASE state OF	
	
0: // IDLE
    Done := FALSE;
    Busy := FALSE;
    Error := FALSE;

    bStopCmd     := FALSE;
    bPowerEnable := TRUE;
    bWriteMode   := FALSE;
    bWait        := FALSE;
    Busy := TRUE;
    state := 10;
    


10: // STOP MOTION
    bStopCmd := TRUE;

    IF fbStopM1.Done AND fbStopM2.Done AND fbStopM3.Done THEN
        bStopCmd := FALSE;
        state := 11;
    END_IF
	
11: // WAIT FOR STANDSTILL
    IF GVL_Axes.Axis1.Status.StandStill 
    AND GVL_Axes.Axis2.Status.StandStill 
    AND GVL_Axes.Axis3.Status.StandStill THEN
        state := 20; // Proceed to Power Off
    END_IF


20: // POWER OFF
    bPowerEnable := FALSE;

    IF NOT fbPowerM1.Status
    AND NOT fbPowerM2.Status
    AND NOT fbPowerM3.Status THEN
        bWait := TRUE;
        state := 30;
    END_IF


30: // WAIT 2s
    IF tWait.Q THEN
        bWait := FALSE;
        state := 40;
    END_IF


40: // WRITE MODE
    bWriteMode := TRUE;

    IF fbWriteModeM1.Done
    AND fbWriteModeM2.Done
    AND fbWriteModeM3.Done THEN
        bWriteMode := FALSE;
        state := 50;
    END_IF

    IF fbWriteModeM1.Error
    OR fbWriteModeM2.Error
    OR fbWriteModeM3.Error THEN
		bWriteMode := FALSE;
        Error := TRUE;
        state := 100;
		Testii := 11;
		 LastErrorCode := fbWriteModeM1.ErrorID;  
    END_IF


50: // POWER ON
   // bPowerEnable := TRUE;
    state := 60;


60: // DONE
    bReadMode := TRUE;

    IF fbReadModeM1.Done
    AND fbReadModeM2.Done
    AND fbReadModeM3.Done THEN

        bReadMode := FALSE;

        IF fbReadModeM1.DriveOperationMode = TO_SINT(TargetMode)
        AND fbReadModeM2.DriveOperationMode = TO_SINT(TargetMode)
        AND fbReadModeM3.DriveOperationMode = TO_SINT(TargetMode) THEN

            Done := TRUE;
            Busy := FALSE;
            state := 0;   // FINISHED SUCCESSFULLY

        ELSE
            Error := TRUE;   // Mode mismatch
            state := 100;
			Testii := 2;
        END_IF
    END_IF

    IF fbReadModeM1.Error
    OR fbReadModeM2.Error
    OR fbReadModeM3.Error THEN
        Error := TRUE;
        state := 100;
		Testii := 3;
	END_IF
	
	100: // Error
		bWriteMode := FALSE;

END_CASE

END_FUNCTION_BLOCK

// ---- POUs/FB_LaunchGame.TcPOU

FUNCTION_BLOCK FB_LaunchGame

VAR_INPUT
    bLaunchSpong       : BOOL;
    bLaunchPeeler      : BOOL;
    bLaunchGoldMiner   : BOOL;
    bLaunchBalloon     : BOOL;
    bLaunchSnowWiper   : BOOL;
    bLaunchSorter      : BOOL;
    bLaunchFlower      : BOOL;
    bLaunchCrazyCar    : BOOL;
END_VAR

VAR_OUTPUT
    eActiveGame : E_GameID := E_GameID.NONE;
    bBusy       : BOOL;
    bError      : BOOL;
END_VAR

VAR
    // Game button rising-edge detection
    trigSpong       : R_TRIG;
    trigPeeler      : R_TRIG;
    trigGoldMiner   : R_TRIG;
    trigBalloon     : R_TRIG;
    trigSnowWiper   : R_TRIG;
    trigSorter      : R_TRIG;
    trigFlower      : R_TRIG;
    trigCrazyCar    : R_TRIG;

    // Windows process launchers
    fbStartProcess : NT_StartProcess;
    fbKillProcess  : NT_StartProcess;

    // Current launch information
    sExePath       : T_MaxString;
    sWorkingDir    : T_MaxString;

    // Requested game information
    eRequestedGame       : E_GameID := E_GameID.NONE;
    sRequestedExePath    : T_MaxString;
    sRequestedWorkingDir : T_MaxString;
    sRequestedExeName    : T_MaxString;

    // Previously launched executable
    sCurrentExeName : T_MaxString;

    // Windows taskkill arguments
    sKillCommand : T_MaxString;

    // One-cycle start signals
    bTriggerStart : BOOL := FALSE;
    bTriggerKill  : BOOL := FALSE;

    // Game switching state
    // 0  = Idle
    // 10 = Issue close request
    // 20 = Wait for close-command acknowledgement
    // 25 = Allow time for process exit
    // 30 = Issue new game launch
    // 40 = Wait for launch acknowledgement
    nState : INT := 0;

    // Wait after Windows accepts close command
    tWaitAfterKill : TON;

    // Diagnostic error code
    nLastProcessErrId : UDINT := 0;
END_VAR


 // ============================================================
 // 1. DETECT HMI BUTTON RISING EDGES
 // ============================================================

trigSpong(CLK := bLaunchSpong);
trigPeeler(CLK := bLaunchPeeler);
trigGoldMiner(CLK := bLaunchGoldMiner);
trigBalloon(CLK := bLaunchBalloon);
trigSnowWiper(CLK := bLaunchSnowWiper);
trigSorter(CLK := bLaunchSorter);
trigFlower(CLK := bLaunchFlower);
trigCrazyCar(CLK := bLaunchCrazyCar);


// ============================================================
// 2. ACCEPT NEW GAME SELECTION ONLY WHEN IDLE
// ============================================================

IF nState = 0 THEN

    IF trigSpong.Q OR
       trigPeeler.Q OR
       trigGoldMiner.Q OR
       trigBalloon.Q OR
       trigSnowWiper.Q OR
       trigSorter.Q OR
       trigFlower.Q OR
       trigCrazyCar.Q THEN

        // ----------------------------------------------------
        // PONG
        // ----------------------------------------------------
        IF trigSpong.Q THEN

            eRequestedGame := E_GameID.PONG;

            sRequestedExePath :=
                'C:\Users\hkhabiri\Desktop\PongV2\RobotGame_BuildV4\Pong.exe';

            sRequestedWorkingDir :=
                'C:\Users\hkhabiri\Desktop\PongV2\RobotGame_BuildV4\';

            sRequestedExeName := 'Pong.exe';


        // ----------------------------------------------------
        // PEELER
        // ----------------------------------------------------
        ELSIF trigPeeler.Q THEN

            eRequestedGame := E_GameID.PEELING;

            sRequestedExePath :=
                'C:\Users\hkhabiri\Desktop\Games\Peeler\EXE_PEELER_2026_10_25\FruitPeeler.exe';

            sRequestedWorkingDir :=
                'C:\Users\hkhabiri\Desktop\Games\Peeler\EXE_PEELER_2026_10_25\';

            sRequestedExeName := 'FruitPeeler.exe';


        // ----------------------------------------------------
        // GOLD MINER
        // ----------------------------------------------------
        ELSIF trigGoldMiner.Q THEN

            eRequestedGame := E_GameID.GOLD_MINER;

            sRequestedExePath :=
                'C:\Users\hkhabiri\Desktop\MotivaGames\GoldMiner\GoldMiner.exe';

            sRequestedWorkingDir :=
                'C:\Users\hkhabiri\Desktop\MotivaGames\GoldMiner\';

            sRequestedExeName := 'GoldMiner.exe';


        // ----------------------------------------------------
        // BALLOON
        // ----------------------------------------------------
        ELSIF trigBalloon.Q THEN

            eRequestedGame := E_GameID.BALLOON;

            sRequestedExePath :=
                'C:\Users\hkhabiri\Desktop\MotivaGames\Balloon\Balloon.exe';

            sRequestedWorkingDir :=
                'C:\Users\hkhabiri\Desktop\MotivaGames\Balloon\';

            sRequestedExeName := 'Balloon.exe';


        // ----------------------------------------------------
        // SNOW WIPER
        // ----------------------------------------------------
        ELSIF trigSnowWiper.Q THEN

            eRequestedGame := E_GameID.SNOW_WIPER;

            sRequestedExePath :=
                'C:\Users\hkhabiri\Desktop\MotivaGames\SnowWiper\SnowWiper.exe';

            sRequestedWorkingDir :=
                'C:\Users\hkhabiri\Desktop\MotivaGames\SnowWiper\';

            sRequestedExeName := 'SnowWiper.exe';


        // ----------------------------------------------------
        // SORTER
        // ----------------------------------------------------
        ELSIF trigSorter.Q THEN

            eRequestedGame := E_GameID.SORTER;

            sRequestedExePath :=
                'C:\Users\hkhabiri\Desktop\Games\Peeler\EXE_Cargo_2026_10_24\Cargo_Sorter_Game.exe';

            sRequestedWorkingDir :=
                'C:\Users\hkhabiri\Desktop\Games\Peeler\EXE_Cargo_2026_10_24\';

            sRequestedExeName := 'Cargo_Sorter_Game.exe';


              // ----------------------------------------------------
        // FLOWER  (= Firefly Garden)
        // ----------------------------------------------------
        ELSIF trigFlower.Q THEN

            eRequestedGame := E_GameID.FLOWER;

            sRequestedExePath :=
                'C:\Users\hkhabiri\Desktop\Games\Peeler\EXE_Firefly_2026_11_06\Firefly Garden Game.exe';

            sRequestedWorkingDir :=
                'C:\Users\hkhabiri\Desktop\Games\Peeler\EXE_Firefly_2026_11_06\';

            sRequestedExeName := 'Firefly Garden Game.exe';



        // ----------------------------------------------------
        // CRAZY CAR
        // ----------------------------------------------------
        ELSIF trigCrazyCar.Q THEN

            eRequestedGame := E_GameID.CRAZY_CAR;

            sRequestedExePath :=
                'C:\Users\hkhabiri\Desktop\Games\SIMON_2\EXE_CrazyCar\CrazyCar.exe';

            sRequestedWorkingDir :=
                'C:\Users\hkhabiri\Desktop\Games\SIMON_2\EXE_CrazyCar\';

            sRequestedExeName := 'CrazyCar.exe';

        END_IF;


        // ----------------------------------------------------
        // BEGIN SWITCH ONLY IF GAME IS DIFFERENT
        // ----------------------------------------------------

        IF eRequestedGame <> eActiveGame THEN

            // Reset launch diagnostics
            bError := FALSE;
            nLastProcessErrId := 0;

            // Disable old game's therapy control
            // during the switching operation
            eActiveGame := E_GameID.NONE;

            // If an old executable is recorded,
            // request its closure first
            IF sCurrentExeName <> '' THEN

                nState := 10;

            ELSE

                // No previous executable recorded
                nState := 30;

            END_IF;

        END_IF;

    END_IF;

END_IF;


// ============================================================
// 3. DEFAULT PROCESS TRIGGERS
//
// Both NT_StartProcess blocks are called every PLC scan.
// START is TRUE for just one PLC scan per request.
// ============================================================

bTriggerKill := FALSE;
bTriggerStart := FALSE;


// ============================================================
// 4. WAIT TIMER
//
// The timer is executed every scan.
// ============================================================

tWaitAfterKill(
    IN := (nState = 25),
    PT := T#1S
);


// ============================================================
// 5. GAME SWITCHING STATE MACHINE
// ============================================================

CASE nState OF

    // --------------------------------------------------------
    // STATE 0: IDLE
    // --------------------------------------------------------
    0:

        // No action


    // --------------------------------------------------------
    // STATE 10: REQUEST CLOSURE OF CURRENT GAME
    // --------------------------------------------------------
    10:

        // Windows taskkill arguments
        // Example:
        // /F /IM "First_Project.exe"

        sKillCommand :=
            CONCAT('/F /IM "', sCurrentExeName);

        sKillCommand :=
            CONCAT(sKillCommand, '"');

        // One-scan rising-edge request
        bTriggerKill := TRUE;

        nState := 20;


    // --------------------------------------------------------
    // STATE 20: WAIT FOR CLOSE COMMAND ACKNOWLEDGEMENT
    // --------------------------------------------------------
    20:

        IF NOT fbKillProcess.BUSY THEN

            IF fbKillProcess.ERR THEN

                // Windows did not accept launch
                // of the taskkill command
                bError := TRUE;

                nLastProcessErrId :=
                    fbKillProcess.ERRID;

                // Do not launch another game
                eRequestedGame := E_GameID.NONE;

                nState := 0;

            ELSE

                // taskkill command was launched
                // Allow time for it to execute
                nState := 25;

            END_IF;

        END_IF;


    // --------------------------------------------------------
    // STATE 25: WAIT AFTER CLOSE REQUEST
    // --------------------------------------------------------
    25:

        IF tWaitAfterKill.Q THEN

            // Previous executable is assumed closed.
            // Actual process exit is NOT verified here.

            sCurrentExeName := '';

            nState := 30;

        END_IF;


    // --------------------------------------------------------
    // STATE 30: REQUEST NEW GAME LAUNCH
    // --------------------------------------------------------
    30:

        sExePath := sRequestedExePath;

        sWorkingDir := sRequestedWorkingDir;

        // One-scan launch request
        bTriggerStart := TRUE;

        nState := 40;


    // --------------------------------------------------------
    // STATE 40: WAIT FOR LAUNCH ACKNOWLEDGEMENT
    // --------------------------------------------------------
    40:

        IF NOT fbStartProcess.BUSY THEN

            IF fbStartProcess.ERR THEN

                bError := TRUE;

                nLastProcessErrId :=
                    fbStartProcess.ERRID;

                eActiveGame := E_GameID.NONE;
                eRequestedGame := E_GameID.NONE;

                nState := 0;

            ELSE

                // Windows accepted the launch command

                eActiveGame := eRequestedGame;

                // Remember current game executable
                // for the next switching operation

                sCurrentExeName :=
                    sRequestedExeName;

                nState := 0;

            END_IF;

        END_IF;

END_CASE;


// ============================================================
// 6. CALL WINDOWS CLOSE COMMAND
//
// Launch taskkill.exe directly, without cmd.exe.
// /F = force process termination
// /IM = executable image name
// ============================================================

fbKillProcess(
    NETID     := '',
    PATHSTR   := 'C:\Windows\System32\taskkill.exe',
    DIRNAME   := 'C:\Windows\System32\',
    COMNDLINE := sKillCommand,
    START     := bTriggerKill,
    TMOUT     := T#5S
);


// ============================================================
// 7. LAUNCH SELECTED UNITY GAME ON MONITOR 3
// ============================================================

fbStartProcess(
    NETID     := '',
    PATHSTR   := sExePath,
    DIRNAME   := sWorkingDir,
    COMNDLINE := '-monitor 2',
    START     := bTriggerStart,
    TMOUT     := T#5S
);


// ============================================================
// 8. MUTUAL EXCLUSION OF ALL HMI GAME BUTTONS
//
// Only the selected game stays TRUE.
// All other GVL_HMI launch flags become FALSE.
// ============================================================

GVL_HMI.bLaunchGameSpongCmd :=
    (eRequestedGame = E_GameID.PONG);

GVL_HMI.bLaunchGamePeelerCmd :=
    (eRequestedGame = E_GameID.PEELING);

GVL_HMI.bLaunchGameGoldMiner :=
    (eRequestedGame = E_GameID.GOLD_MINER);

GVL_HMI.bLaunchGameBalloonAssesment :=
    (eRequestedGame = E_GameID.BALLOON);

GVL_HMI.bLaunchGameSnowWiper :=
    (eRequestedGame = E_GameID.SNOW_WIPER);

GVL_HMI.bLaunchGameSorter :=
    (eRequestedGame = E_GameID.SORTER);

GVL_HMI.bLaunchGameFlower :=
    (eRequestedGame = E_GameID.FLOWER);

GVL_HMI.bLaunchGameCrazyCar :=
    (eRequestedGame = E_GameID.CRAZY_CAR);


// ============================================================
// 9. PROCESS STATUS
// ============================================================

bBusy :=
    (nState <> 0)
    OR fbStartProcess.BUSY
    OR fbKillProcess.BUSY;

END_FUNCTION_BLOCK

// ---- POUs/Sorter Game/FB_SorterGame.TcPOU
FUNCTION_BLOCK FB_SorterGame
VAR_INPUT
    bEnable                   : BOOL;
    stCartesianPosePercentage : ST_CartesianPose;  // same as PeelingGame
	CartesianForcefx            : LREAL ; 
  //  RehabilitationController: E_ControllerType;
	CartesianVx : LREAL;
END_VAR
VAR
    stToUnity : ST_SorterToUnity;
	stFromUnity : ST_UnityToSorter;
	FXThreshold    : REAL := 3.0 ;  // Minimum Force to create Resistive Force;
	VXThreshold : LREAL := 10.0;
END_VAR

VAR_OUTPUT
	stJointTargetTorque : ST_JointTorque;
END_VAR

// Default outputs
stJointTargetTorque.M1 := 0.0;
stJointTargetTorque.M2 := 0.0;
stJointTargetTorque.M3 := 0.0;

stToUnity.GameIsActive := FALSE;


IF bEnable THEN

    // Send X position to Unity
    stToUnity.fX := stCartesianPosePercentage.X;

    IF NOT stFromUnity.bGameClosed THEN

        stToUnity.GameIsActive := TRUE;


        (****************************************************
            CONDITION 1: POSITIVE X MOVEMENT

            Both Vx and Fx must be positive
            and exceed their thresholds.

            Apply NEGATIVE resistance.
        *****************************************************)

